# B&R Automation Studio project Palletizer_Final_project_2
Automation Studio 4.10.2.37

## Configuration Config1

### Hardware
```
4PP065_0351_P74 : 4PP065.0351-P74 v1.0.4.0
  Connector IF5:
    ActivateDevice = 1
    Mode = Manual
    InternetAddress = 127.0.0.1
    Vnc1
    VncVcObjectName1 = Visu_R
    VncKeyMappingFile1 = VC\PS2-Keyboard.dis
    VncAuthentication1 = 1
    VncPasswordViewOnly1 = r
    VncPasswordViewControl1 = w
  ConfigurationID = Palletizer_Final_project_Config1
  Simulation = 1
  FileDevice1
  FileDeviceName1 = USER
  FileDevicePath1 = USER_PATH
  KeyMappingFile = VC\4PP065_0351_P74.dis
```

## Logical view

Binary libraries used (declarations not repeated): operator, runtime, astime, AsIecCon, AsTCP, standard, AsArLog, AsBrStr

### Global.var - Global variables
```iecst
(*FEEDERSTATION*)
(*Insert your comment here.*)
VAR
	OperationType : INT;
	ENABLE_CONVEYER_END : BOOL;
	ENABLE_CONVEYER_TURN1 : BOOL;
	TURNPUSHER_FAULT : BOOL;
	ENABLE_TURNPUSHER : BOOL;
	DISABLE_TURNPUSHER : BOOL;
	TURNPUSHER_ENABLED : BOOL;
	TURNPUSHER_DISABLED : BOOL;
	PUSHER_FAULT : BOOL;
	ENABLE_PUSHER : BOOL;
	PUSHER_DISABLED : BOOL;
	PUSHER_ENABLED : BOOL;
	ENABLE_CONVEYOR_IF : BOOL;
	START_FEEDER : BOOL;
	LASER_SENSOR_IR : BOOL;
	FIRST_LAYER_OPERATION : BOOL;
	NUM_BOX_COUNTED : INT;
	COUNT_LASER_SENSOR_IR : INT;
	LASER_SENSOR_2_IR : BOOL;
	ACTUAL_BOXES : INT;
	ACTUAL_CARRIAGE_POS : REAL;
	CARRIAGE_TRG_POS : REAL;
	CARRIAGE_RCHD_POS : BOOL;
	SIMULATE_FAULT_CARRIAGE_2 : BOOL;
	FEERDER_BOXES_DELIVERED : BOOL;
	START_AGAIN_FEEDER : BOOL;
	FEEDER_EMERGENCY_STOP : BOOL;
	FEEDER_IMMEDIATE_STOP : BOOL;
	FEEDER_ON_PHASE_STOP : BOOL;
	FEEDER_ON_PHASE_STOP_WAIT : BOOL;
	ENABLE_SLIDE_RAIL_RIGHT : BOOL;
	VACUUM_BOX_CRANE_ENABLED : BOOL;
	ENABLE_VACUUM_BOX_CRANE : BOOL;
	VACUUM_BOX_CRANE_FAULT : BOOL;
	ENABLE_PUSHER_X : BOOL;
	ENABLE_PUSHER_Z : BOOL;
	ENABLE_CARTBORAD : BOOL;
	GANTRY_CRANE_RCHD_POS : BOOL;
	FAULT_GANTRY_CRANE : BOOL;
	ACTUAL_GANTRY_CRANE_POS : REAL;
	GANTRY_CRANE_TRG_POS : REAL;
	BOX_CRANE_RCHD_POS : BOOL;
	FAULT_BOX_CRANE : BOOL;
	ACTUAL_BOX_CRANE_POS : REAL;
	BOX_CRANE_TRG_POS : REAL;
	START_CRANE : BOOL;
	CRANE_WAIT_BOXES : BOOL;
	SECOND_LAYER_OPERATION : BOOL;
	LASER_SENSOR_IR_MEM : BOOL;
	LASER_SENSOR_2_IR_MEM : BOOL;
	CRANE_ON_PHASE_STOP : BOOL;
	CRANE_ON_PHASE_STOP_WAIT : BOOL;
	CRANE_EMERGENCY_STOP : BOOL;
	CRANE_IMMEDIATE_STOP : BOOL;
	FAULT_PALLET_CONVEYOR_2 : BOOL;
	PALLET_CONVEYOR_2_TRG_VEL : REAL;
	PALLET_LIFTER_RCHD_POS : BOOL;
	FAULT_PALLET_LIFTER : BOOL;
	ACTUAL_PALLET_LIFTER_POS : REAL;
	PALLET_LIFTER_TRG_POS : REAL;
	PALLET_FORK_ENABLED : BOOL;
	ENABLE_PALLET_FORK : BOOL;
	PALLET_FORK_FAULT : BOOL;
	ENABLE_PALLET_CONVEYOR_1 : BOOL;
	PALLET_CONVEYOR_1_FAULT : BOOL;
	PALLET_LIGHT_BARRIER_2 : BOOL;
	PALLET_LIGHT_BARRIER_1 : BOOL;
	PALLET_WAIT_BOXES : BOOL;
	AFTER_IMMEDIATE_STOP : BOOL; (*gives acces to the pallet state after the immediate stop*)
	START_PALLET : BOOL;
	PALLET_ON_PHASE_STOP_WAIT : BOOL;
	PALLET_EMERGENCY_STOP : BOOL;
	PALLET_IMMEDIATE_STOP : BOOL;
	PALLET_ON_PHASE_STOP : BOOL;
	BUTTON_START : BOOL;
	BUTTON_STOP : BOOL;
	BUTTON_EMERGENCY_STOP : BOOL;
	BUTTON_IMMEDIATE_STOP : BOOL;
	BUTTON_ON_PHASE_STOP : BOOL;
	BUTTON_INITIALIZATION : BOOL;
	blink_start : BOOL;
	blink_stop : BOOL;
	blink_ermergency : BOOL;
	blink_immediatestop : BOOL;
	blink_onphasestop : BOOL;
	blink_Fauld : BOOL;
	FEERDER_WAIT_TO_DELIVER_BOXES : BOOL;
	CRANE_BOXES_DELIVERED : BOOL;
	CARRIAGE_2_FAULT : BOOL;
	CONVEYOR_IF_FAULT : BOOL;
	SIMULATE_FAULT_PUSHER : BOOL;
	SIMULATE_FAULT_TURNPUSHER : BOOL;
	SIMULATE_FAULT_GANTRY_CRANE : BOOL;
	GANTRY_CRANE_FAULT : BOOL;
	SIMULATE_FAULT_BOX_CRANE : BOOL;
	BOX_CRANE_FAULT : BOOL;
	SIMULATE_FAULT_SLIDE_RIGTH : BOOL;
	SIMULATE_FAULT_SLIDE_RAIL_RIGHT : BOOL;
	SLIDE_RAIL_RIGHT_FAULT : BOOL;
	SIMULATE_FAULT_VACUUM_BOX_CRANE : BOOL;
	SIMULATE_FAULT_PUSHER_X : BOOL;
	PUSHER_X_FAULT : BOOL;
	SIMULATE_FAULT_PUSHER_Z : BOOL;
	PUSHER_Z_FAULT : BOOL;
	SIMULATE_FAULT_CARTBORAD : BOOL;
	CARTBORAD_FAULT : BOOL;
	SIMULATE_FAULT_PALLET_LIFTER : BOOL;
	PALLET_LIFTER_FAULT : BOOL;
	SIMULATE_FAULT_PALLET_CONVEYOR_2 : BOOL;
	PALLET_CONVEYOR_2_FAULT : BOOL;
	SIMULATE_FAULT_PALLET_FORK : BOOL;
	ENABLE_CONVEYOR_TURN1 : BOOL;
	CONVEYOR_TURN1_FAULT : BOOL;
	ENABLE_CONVEYOR_END : BOOL;
	CONVEYOR_END_FAULT : BOOL;
	LED_ALARM_INFORMATION : BOOL;
	LED_ALARM_ANOMALY : BOOL;
	LED_ALARM_ALARM : BOOL;
	LED_ALARM_WARNING : BOOL;
	SM_ON_PHASE_STOP : BOOL;
	SM_IMMEDIATE_STOP : BOOL;
	SM_EMERGENCY_STOP : BOOL;
	SM_IMMEDIATE_STOP_CAT1 : BOOL;
	SM_IMMEDIATE_STOP_CAT2 : BOOL;
	SM_IMMEDIATE_STOP_CAT3 : BOOL;
	LED_MATERIALS_RUN_OUT : BOOL;
	SM_ON_PHASE_STOP_CAT2 : BOOL;
	SM_ON_PHASE_STOP_CAT1 : BOOL;
	PALLET_ON_PHASE_STOP_REMOVE : BOOL;
	SM_ON_PHASE_STOP_CAT_2 : BOOL;
	boxcrane_Cartboard_ALMOST_FINISH : BOOL;
	boxcrane_Cartboard_FINISH : BOOL;
	pallet_lifter_ALMOST_FINISH : BOOL;
	pallet_lifter_FINISH : BOOL;
	POWER_ON_FEEDER : BOOL;
	POWER_ON_CRANE : BOOL;
	POWER_ON_PALLET : BOOL;
	POWER_MACHINE : BOOL;
	POWER_ON_BUTTON : BOOL;
	PALLET_ON_PHASE_STOP_IDLE : BOOL;
	COUNT_PALLET_NUMBER : INT := 5;
	COUNT_CARTBOARD_NUMBER : INT := 25;
	COUNT_BOXES_NUMBER : INT;
	blink_emergencvy_stop : BOOL;
	blink_immediate_stop : BOOL;
	blink_OnPhase_stop : BOOL;
	PALLET_STOP : BOOL;
	CRANE_STOP : BOOL;
	FEEDER_STOP : BOOL;
END_VAR
```

### MNG_Package.var
```iecst
(*                                                                            *)
(* File generated by the B&R AS 4 control config generator                    *)
(*                                                                            *)
(*     Provider: machineering                                                 *)
(*  Application: industrialPhysics_2.4.master                                 *)
(* Architecture: Windows 64 Bit                                               *)
(*      Version: 2.4.10491.master                                             *)
(*        Build: 164f85bec                                                    *)
(*         Date: 2020-05-19, Time: 12:11:21                                   *)
(*                                                                            *)
VAR
	ComTCP_SimInputs : ComTCP_INPUTS_32BIT := (0);
	ComTCP_SimOutputs : ComTCP_OUTPUTS_32BIT := (0);
	ComTCP_SimServerAddress : STRING[15] := '127.0.0.1';
	ComTCP_SimServerPort : UINT := 5000;
	ComTCP_SimSendCycleTime : TIME := T#5ms;
	ComTCP_SimActive : BOOL := FALSE;
END_VAR
```

### MNG_Package.typ
```iecst
(*                                                                            *)
(* File generated by the B&R AS 4 control config generator                    *)
(*                                                                            *)
(*     Provider: machineering                                                 *)
(*  Application: industrialPhysics_2.4.master                                 *)
(* Architecture: Windows 64 Bit                                               *)
(*      Version: 2.4.10491.master                                             *)
(*        Build: 164f85bec                                                    *)
(*         Date: 2020-05-19, Time: 12:11:21                                   *)
(*                                                                            *)

TYPE
	ComTCP_INPUTS_32BIT : 	STRUCT
		NumSignals : INT := 15;
		laser_sensor_IR : BOOL := 0; (* BOOL laser_sensor_IR *)
		laser_sensor2_IR : BOOL := 0; (* BOOL laser_sensor2_IR *)
		carriage_2_AXIS : REAL := 0.0; (* REAL carriage_2_AXIS *)
		carriage_2_RCHD : BOOL := 0; (* BOOL carriage_2_RCHD *)
		turnpusher_LBK : BOOL := 0; (* BOOL turnpusher_LBK *)
		turnpusher_LFR : BOOL := 0; (* BOOL turnpusher_LFR *)
		gantry_crane_AXIS : REAL := 0.0; (* REAL gantry_crane_AXIS *)
		box_crane_AXIS : REAL := 0.0; (* REAL box_crane_AXIS *)
		vaccum_box_crane_VACUUM : BOOL := 0; (* BOOL vaccum_box_crane_VACUUM *)
		pallet_light_barrier_1_IR : BOOL := 0; (* BOOL pallet_light_barrier_1_IR *)
		pallet_light_barrier_2_IR : BOOL := 0; (* BOOL pallet_light_barrier_2_IR *)
		pusher_LBK : BOOL := 0; (* BOOL pusher_LBK *)
		pusher_LFR : BOOL := 0; (* BOOL pusher_LFR *)
		pallet_lifter_AXIS : REAL := 0.0; (* REAL pallet_lifter_AXIS *)
		pallet_fork_left_FB : BOOL := 0; (* BOOL pallet_fork_left_FB *)
	END_STRUCT;
	ComTCP_OUTPUTS_32BIT : 	STRUCT
		NumSignals : INT := 18;
		cartboard_TRIG : BOOL := 0; (* BOOL cartboard_TRIG *)
		conveyor_if_FWD : BOOL := 0; (* BOOL conveyor_if_FWD *)
		conveyer_turn1_FWD : BOOL := 0; (* BOOL conveyer_turn1_FWD *)
		conveyer_end_FWD : BOOL := 0; (* BOOL conveyer_end_FWD *)
		carriage_2_TGT_POS : REAL := 0.0; (* REAL carriage_2_TGT_POS *)
		turnpusher_FWD : BOOL := 0; (* BOOL turnpusher_FWD *)
		turnpusher_BWD : BOOL := 0; (* BOOL turnpusher_BWD *)
		gantry_crane_TGT_POS : REAL := 0.0; (* REAL gantry_crane_TGT_POS *)
		box_crane_TGT_POS : REAL := 0.0; (* REAL box_crane_TGT_POS *)
		slide_rail_right_EN : BOOL := 0; (* BOOL slide_rail_right_EN *)
		vaccum_box_crane_GRIP : BOOL := 0; (* BOOL vaccum_box_crane_GRIP *)
		pusher_z_EN : BOOL := 0; (* BOOL pusher_z_EN *)
		pusher_x_EN : BOOL := 0; (* BOOL pusher_x_EN *)
		pallet_conveyor_2_ACT_VEL : REAL := 0.0; (* REAL pallet_conveyor_2_ACT_VEL *)
		pusher_FW : BOOL := 0; (* BOOL pusher_FW *)
		pallet_lifter_TGT_POS : REAL := 0.0; (* REAL pallet_lifter_TGT_POS *)
		pallet_fork_left_EN : BOOL := 0; (* BOOL pallet_fork_left_EN *)
		pallet_conveyor_1_FWD : BOOL := 0; (* BOOL pallet_conveyor_1_FWD *)
	END_STRUCT;
END_TYPE
```

### Package Logical/Libraries - Global libraries

### Library Logical/Libraries/G_Device (IEC)

#### Types.typ - Exported data types
```iecst
TYPE
	DeviceStateType :
	(
		DeviceEnabledState		:=2,
		DeviceEnablePhaseState	:=1,
		DeviceDisabledState		:=0,
		DeviceDisablePhaseState	:=3
	);
END_TYPE
```

#### Constants.var - Exported constants
```iecst
VAR CONSTANT
	DEVICE_ACTUATION_MASK : INT := 2#00001111;
	DEVICE_FEEDBACK_MASK : INT := 2#11110000;
	DEVICE_WITH_ENABLE_FEEDBACK : INT := 2#00010000;
	DEVICE_WITH_DISABLE_FEEDBACK : INT := 2#00100000;
	DEVICE_WITHOUT_FEEDBACK : INT := 2#01000000;
	DEVICE_WITH_SINGLE_ACTUATION : INT := 2#00000001;
	DEVICE_WITH_DOUBLE_ACTUATION : INT := 2#00000011;
	DEVICE_WITH_DA_NO_RETAIN : INT := 2#00000010;
	DEVICE_WITH_DOUBLE_FEEDBACK : INT := 2#00110000;
END_VAR
```

#### G_Device.fun - Exported functions and function blocks
```iecst
{REDUND_ERROR} FUNCTION_BLOCK Generic_Device (*TODO: Add your comment here*) (*$GROUP=User,$CAT=User,$GROUPICON=User.png,$CATICON=User.png*)
	VAR_INPUT
		DeviceClock : {REDUND_UNREPLICABLE} BOOL;
		DeviceDisabledSensor : {REDUND_UNREPLICABLE} BOOL;
		DeviceEnabledSensor : {REDUND_UNREPLICABLE} BOOL;
		DeviceEnabled : {REDUND_UNREPLICABLE} BOOL;
		DeviceDisabled : {REDUND_UNREPLICABLE} BOOL;
		DeviceType : {REDUND_UNREPLICABLE} INT;
		DeviceOperation : {REDUND_UNREPLICABLE} INT;
		DeviceEnablePreset : {REDUND_UNREPLICABLE} BOOL;
		DeviceEnableTime : {REDUND_UNREPLICABLE} INT;
		DeviceDisableTime : {REDUND_UNREPLICABLE} INT;
		DeviceDiagnosticsEnabled : BOOL;
		SimulationDeviceFault : BOOL;
	END_VAR
	VAR_OUTPUT
		EnableDevice : {REDUND_UNREPLICABLE} BOOL;
		DeviceNotInitialized : {REDUND_UNREPLICABLE} BOOL;
		DisableDevice : {REDUND_UNREPLICABLE} BOOL;
		DeviceDisabledSensorFault : {REDUND_UNREPLICABLE} BOOL;
		DeviceEnabledSensorFault : {REDUND_UNREPLICABLE} BOOL;
		DeviceActuatorFault : {REDUND_UNREPLICABLE} BOOL;
		DeviceFault : {REDUND_UNREPLICABLE} BOOL;
	END_VAR
	VAR_IN_OUT
		DeviceEnableRequest : BOOL;
		DeviceDisableRequest : BOOL;
	END_VAR
	VAR
		DeviceTimer : {REDUND_UNREPLICABLE} INT;
	END_VAR
	VAR RETAIN
		DeviceState : {REDUND_UNREPLICABLE} DeviceStateType;
	END_VAR
	VAR
		Timeout : {REDUND_UNREPLICABLE} BOOL := FALSE;
	END_VAR
	VAR CONSTANT
		INIT : INT := 0;
	END_VAR
	VAR
		WaitNominalStateCounter : INT := 20;
		SimulationDeviceActuatorFault : BOOL;
	END_VAR
END_FUNCTION_BLOCK
```

#### Generic_Device.st
```iecst
(* TODO: Add your comment here *)
FUNCTION_BLOCK Generic_Device

	//I-) DEVICE CLOCK HANDLER
	IF (DeviceClock AND (DeviceTimer > 0))THEN
		DeviceTimer := DeviceTimer - 1;
		WaitNominalStateCounter := WaitNominalStateCounter	- 1;
	END_IF;

	//II-) DEVICE SENSORS HANDLER
	CASE (DeviceType AND DEVICE_FEEDBACK_MASK) OF

		DEVICE_WITH_ENABLE_FEEDBACK:

			DeviceDisabledSensor := NOT DeviceEnabledSensor AND
			((DeviceState = DeviceDisabledState) OR (DeviceState = DeviceDisablePhaseState AND Timeout));
			//Pre-elaborations actuators
			DeviceDisabled := NOT DeviceEnabled AND ((DeviceState = DeviceDisabledState) OR
			(DeviceState = DeviceDisablePhaseState AND Timeout));

		DEVICE_WITH_DISABLE_FEEDBACK :

			DeviceEnabledSensor := NOT DeviceDisabledSensor AND
			((DeviceState = DeviceEnabledState) OR (DeviceState = DeviceEnablePhaseState AND Timeout));
			//Pre-elaborations actuators
			DeviceEnabled := NOT DeviceDisabled AND ((DeviceState = DeviceEnabledState) OR
			(DeviceState = DeviceEnablePhaseState AND Timeout));

		DEVICE_WITHOUT_FEEDBACK:

			DeviceEnabledSensor := (DeviceState = DeviceEnabledState) OR ((DeviceState = DeviceEnablePhaseState) AND Timeout);
			DeviceDisabledSensor := (DeviceState = DeviceDisabledState) OR ((DeviceState = DeviceDisablePhaseState) AND Timeout);
			//Pre-elaborations actuators
			DeviceEnabled := (DeviceState = DeviceEnabledState) OR (DeviceState = DeviceEnablePhaseState AND Timeout);
			DeviceDisabled := (DeviceState = DeviceDisabledState) OR (DeviceState = DeviceDisablePhaseState AND Timeout);

	END_CASE;

	//III-) DEVICE INITIALIZATION HANDLER
	IF (DeviceOperation = INIT) THEN
		// Device sensor handler
		CASE (DeviceType AND DEVICE_FEEDBACK_MASK) OF

			DEVICE_WITH_ENABLE_FEEDBACK:
				DeviceDisabled := NOT DeviceEnabled;

			DEVICE_WITH_DISABLE_FEEDBACK :
				DeviceEnabled := NOT DeviceDisabled;

			DEVICE_WITHOUT_FEEDBACK:
				DeviceEnabled := DeviceEnablePreset;
				DeviceDisabled := NOT DeviceEnabled;

		END_CASE;

		DeviceEnableRequest := FALSE;
		DeviceDisableRequest := FALSE;

		IF (DeviceEnablePreset) THEN
			EnableDevice := TRUE;
			DeviceTimer := DeviceEnableTime;
			IF (NOT (DeviceDisabled AND DeviceEnabled)) THEN
				DeviceState := DeviceEnablePhaseState;
			ELSE
				DeviceState := DeviceEnabledState;
			END_IF;
			DeviceNotInitialized := NOT DeviceEnabled OR DeviceDisabled;
		ELSE
			EnableDevice := FALSE;
			DeviceTimer := DeviceDisableTime;
			IF (NOT (DeviceDisabled AND DeviceEnabled)) THEN
				DeviceState := DeviceDisablePhaseState;
			ELSE
				DeviceState := DeviceDisabledState;
			END_IF;
			DeviceNotInitialized := (DeviceEnabled OR NOT DeviceDisabled);
		END_IF;
	END_IF;

	IF NOT SimulationDeviceFault THEN
		//IV-) DEVICE CONTROL HANDLER (GENERIC DEVICE FSM IMPLEMENTATION)
		CASE (DeviceState) OF

			DeviceDisabledState:
				DeviceDisableRequest := FALSE;
				IF (DeviceEnableRequest) THEN
					EnableDevice := TRUE;
					DeviceTimer := DeviceEnableTime;
					DeviceState := DeviceEnablePhaseState;
				END_IF;

			DeviceEnablePhaseState:
				IF DeviceDisableRequest THEN
					DeviceEnableRequest	:= FALSE;
					EnableDevice	:= FALSE;
					DeviceTimer	:= DeviceDisableTime;
					DeviceState	:= DeviceDisablePhaseState;
				END_IF;
				IF DeviceEnabledSensor THEN
					DeviceEnableRequest := FALSE;
					DeviceTimer	:= 0;
					DeviceState := DeviceEnabledState;
				END_IF;

			DeviceEnabledState:
				DeviceEnableRequest	:= FALSE;
				IF DeviceDisableRequest THEN
					EnableDevice := FALSE;
					DeviceTimer	:= DeviceDisableTime;
					DeviceState := DeviceDisablePhaseState;
				END_IF;

			DeviceDisablePhaseState:
				IF DeviceEnableRequest THEN
					DeviceDisableRequest	:= FALSE;
					EnableDevice	:= TRUE;
					DeviceTimer	:= DeviceEnableTime;
					DeviceState	:= DeviceEnablePhaseState;
				END_IF;

				IF DeviceDisabledSensor THEN
					DeviceDisableRequest := FALSE;
					DeviceTimer	:= 0;
					DeviceState := DeviceDisabledState;
				END_IF;

		END_CASE;

	END_IF;

	//handler timer
	IF (DeviceTimer = 0) THEN
		Timeout := TRUE ;

	ELSE
		Timeout := FALSE ;

	END_IF;

	//V-) DEVICE DIAGNOSTICS HANDLER (GENERATION OF DIAGNOSIS INFORMATION),
	DeviceDisabledSensorFault := (( NOT EnableDevice AND NOT DeviceDisabledSensor AND NOT DeviceEnabledSensor) OR (EnableDevice AND DeviceDisabledSensor AND DeviceEnabledSensor)) AND Timeout;

	DeviceEnabledSensorFault := ((NOT EnableDevice AND DeviceDisabledSensor AND DeviceEnabledSensor) OR (EnableDevice AND NOT DeviceDisabledSensor AND NOT DeviceEnabledSensor)) AND Timeout;

	DeviceActuatorFault := ((NOT EnableDevice AND NOT DeviceDisabledSensor AND DeviceEnabledSensor AND Timeout) OR (EnableDevice AND DeviceDisabledSensor AND NOT DeviceEnabledSensor AND Timeout)) AND Timeout;
	//DeviceActuatorFault

	DeviceFault :=	DeviceDisabledSensorFault OR DeviceEnabledSensorFault OR SimulationDeviceFault ;

	//VI-) DEVICE ACTUATORS HANDLER (Post-elaborations actustors)
	IF (DeviceType AND DEVICE_ACTUATION_MASK)= DEVICE_WITH_SINGLE_ACTUATION THEN
		//Nothing to do, just use EnableDevice
	END_IF;
	IF	(DeviceType AND DEVICE_ACTUATION_MASK)= DEVICE_WITH_DOUBLE_ACTUATION THEN
		DisableDevice := NOT EnableDevice;
	END_IF;
	IF	(DeviceType AND DEVICE_ACTUATION_MASK)= DEVICE_WITH_DA_NO_RETAIN THEN
		EnableDevice := EnableDevice AND (DeviceState = DeviceEnablePhaseState);
		DisableDevice := NOT EnableDevice AND (DeviceState = DeviceDisablePhaseState);
	END_IF;
	IF	DeviceActuatorFault AND (DeviceTimer = 0) AND WaitNominalStateCounter = 0  THEN

		SimulationDeviceActuatorFault := TRUE;
		WaitNominalStateCounter := 20;

	ELSE
		SimulationDeviceActuatorFault := FALSE;
	END_IF;

END_FUNCTION_BLOCK
```

### Library Logical/Libraries/G_Axis (IEC)

#### Types.typ - Exported data types
```iecst
TYPE

	GenericAxisType :
		(
		WaitpowerON,
		WaitHoming,
		CheckCommand,
		WaitPowerOFF,
		WaitStop,
		WaitMoveTRG_POS,
		ErrorState,
		WaitMoveTRG_VEL

	);

END_TYPE
```

#### Constants.var - Exported constants
```iecst
VAR CONSTANT
	POWEROFF : DWORD := 1;
	STOP : DWORD := 2;
	HOMING : DWORD := 3;
	TARGETPOSITION : DWORD := 4;
	Notbusy : DWORD := 0;
	TARGETVELOCITY : DWORD := 5;
END_VAR
```

#### G_Axis.fun - Exported functions and function blocks
```iecst
{REDUND_ERROR} FUNCTION_BLOCK Generic_Axis (*TODO: Add your comment here*) (*$GROUP=User,$CAT=User,$GROUPICON=User.png,$CATICON=User.png*)
	VAR_INPUT
		PowerON : BOOL;
		DeviceTimer : INT;
		Actual_position : REAL;
		Input_Target_Position : REAL;
		Reached_Postion : BOOL;
		InputSimulateError : BOOL;
		Actual_Command : DWORD;
		DeviceClock : BOOL;
		DeviceFeedback : BOOL;
	END_VAR
	VAR_OUTPUT
		Powered : BOOL;
		Output_Target_Position : REAL;
		InPosition : BOOL;
		InVelocity : BOOL;
		OutputSimulateError : BOOL;
	END_VAR
	VAR
		Generic_Axis_State : GenericAxisType;
		Timer : INT;
		TimeOut : BOOL;
	END_VAR
	VAR_INPUT
		Input_Target_Velocity : REAL;
	END_VAR
	VAR_OUTPUT
		Output_Target_Velocity : REAL;
	END_VAR
END_FUNCTION_BLOCK
```

#### Generic_Axis.st
```iecst
(* TODO: Add your comment here *)
FUNCTION_BLOCK Generic_Axis
	IF (DeviceClock AND (Timer > 0))THEN
		Timer := Timer - 1;

		END_IF;

	CASE Generic_Axis_State OF

		WaitpowerON:
			IF PowerON THEN
				//all output false
				Powered:= FALSE;
				InPosition	:= FALSE;
				InVelocity	:= FALSE;
				Timer		:= DeviceTimer;
	  			Generic_Axis_State:=WaitHoming;
			END_IF;
		WaitHoming:

			IF TimeOut THEN
				Powered:= TRUE;
				TimeOut		:= FALSE;
				Output_Target_Position:=0.0;
				Output_Target_Velocity:=0.0;
				Actual_Command := Notbusy;
				IF NOT PowerON THEN
					Generic_Axis_State:= WaitpowerON;
				ELSE
					IF Actual_position=0.0 THEN
						InPosition	:= TRUE;
						InVelocity	:= FALSE;
						Generic_Axis_State:= CheckCommand;
					END_IF;
				END_IF;
			END_IF;
		CheckCommand:
			IF Actual_Command = POWEROFF  THEN
				Actual_Command := Notbusy;
				Generic_Axis_State:= WaitPowerOFF;
			END_IF;
			IF Actual_Command = STOP THEN
				Actual_Command := Notbusy;
				Generic_Axis_State:= WaitStop;
			END_IF;
			IF Actual_Command = HOMING THEN
				Actual_Command := Notbusy;
				InVelocity	:= TRUE;
				Generic_Axis_State:= WaitHoming;
			END_IF;
			IF Actual_Command = TARGETPOSITION THEN
				Actual_Command := Notbusy;
				IF Input_Target_Position <> Actual_position THEN
					InVelocity	:= TRUE;
					Timer		:= DeviceTimer;
	  				Generic_Axis_State:= WaitMoveTRG_POS;
				ELSE
					Generic_Axis_State:= CheckCommand;
				END_IF;
			END_IF;
			InPosition	:= FALSE;
			IF Actual_Command = TARGETVELOCITY THEN
				Actual_Command := Notbusy;
				IF Input_Target_Velocity <> Output_Target_Velocity THEN
					InVelocity	:= TRUE;
					Timer		:= DeviceTimer;
					Generic_Axis_State:= WaitMoveTRG_VEL;
				ELSE
					Generic_Axis_State:= CheckCommand;
				END_IF;
			END_IF;
		WaitPowerOFF:
			PowerON := FALSE;
			InPosition	:= FALSE;
			InVelocity	:= FALSE;
			Generic_Axis_State:=WaitHoming;
		WaitStop:

			IF InVelocity THEN
		  		Output_Target_Position:=Actual_position + 0.1; //bias link to the dealy
				IF Reached_Postion THEN

		  			InPosition	:= FALSE;
					InVelocity	:= FALSE;
				END_IF;
			END_IF;
			IF OutputSimulateError THEN
				Generic_Axis_State:= ErrorState;
			ELSE
				Generic_Axis_State:= CheckCommand;
			END_IF;

		WaitMoveTRG_POS:
			Output_Target_Position := Input_Target_Position;
			IF TimeOut THEN
				IF DeviceFeedback AND Reached_Postion THEN
					InPosition	:= TRUE;
					InVelocity	:= FALSE;
					TimeOut		:= FALSE;
					Generic_Axis_State:= CheckCommand;
				END_IF;

				IF NOT DeviceFeedback AND (Input_Target_Position = Actual_position)	 THEN
					InPosition	:= TRUE;
					InVelocity	:= FALSE;
					TimeOut		:= FALSE;
					Generic_Axis_State:= CheckCommand;
				END_IF;

			END_IF;
		WaitMoveTRG_VEL:
			Output_Target_Velocity := Input_Target_Velocity;
			IF TimeOut THEN
				IF NOT DeviceFeedback THEN
					TimeOut		:= FALSE;
					Generic_Axis_State:= CheckCommand;
				END_IF;
			END_IF;

		ErrorState:
			IF NOT InputSimulateError THEN //wait for the Simulated Error to be set back
				OutputSimulateError:=FALSE;
			Generic_Axis_State:= WaitHoming;
			END_IF;

	END_CASE;
	IF Timer=0 THEN
		TimeOut	:= TRUE;
	END_IF;
	IF InputSimulateError THEN
		OutputSimulateError:=TRUE;
		Generic_Axis_State:= WaitStop;
	END_IF;

END_FUNCTION_BLOCK
```

### Library Logical/Libraries/G_SM (IEC)

#### Constants.var - Exported constants
```iecst
VAR CONSTANT
	SIGNAL_TYPE_MASK : INT := 2#00000111;
	ALARM : INT := 2#00000001;
	ANOMALY : INT := 2#00000010;
	WARNING : INT := 2#00000011;
	INFORMATION : INT := 2#00000100;
	AUX_RESET : INT := 2#10100000;
	AUTO_CONDITIONED_RESET : INT := 2#01100000;
	NONE : DWORD := 16#0000;
	INIT : INT := 0;
	RUN : INT := 1;
	START_CONFIGURATION : INT := 2;
	CONFIGURATION : INT := 3;
	START_GENERATION : INT := 4;
	GENERATION : INT := 5;
	EMERGENCY_STOP : DWORD := 16#0001;
	IMMEDIATE_STOP : DWORD := 16#0002;
	ON_PHASE_STOP : DWORD := 16#0004;
	MATERIALS_RUN_OUT_LAMP : DWORD := 16#0006;
	MATERIALS_RUN_OUT_BUZZER : DWORD := 16#0008;
END_VAR
```

#### G_SM.fun - Exported functions and function blocks
```iecst
{REDUND_ERROR} FUNCTION_BLOCK GenericSignalHandler (*TODO: Add your comment here*) (*$GROUP=User,$CAT=User,$GROUPICON=User.png,$CATICON=User.png*)
	VAR_INPUT
		OperationType : INT;
		SignalType : DINT;
		Reset : BOOL;
		KeyReset : BOOL;
		ActivationSignal : BOOL;
		SignalCode : INT;
		SignalOutput : DWORD;
		CondKeyReset : BOOL;
	END_VAR
	VAR_OUTPUT
		NumberOfAlarms : INT;
		NumberOfAnomalies : INT;
		NumberOfWarnings : INT;
		NumberOfInformation : INT;
		ResetEnable : BOOL;
		SignalOutputs : DWORD;
		NumberOfActiveAlarms : INT;
		NumberOfActiveAnomalies : INT := 0;
		NumberOfActiveWarning : INT;
		NumberOfActiveInformation : INT;
		ActiveSignalCodes : ARRAY[0..24] OF INT;
		AuxResetEnable : BOOL;
		AutoCondResetEnable : BOOL;
		LedSignalInformation : BOOL;
		LedSignalAnomaly : BOOL;
		LedSignalWarning : BOOL;
		LedSignalAlarm : BOOL;
		MySignalCode : INT;
	END_VAR
	VAR
		ResetActivation : BOOL;
		ResetOld : BOOL;
		KeyResetOld : BOOL;
		Index : INT;
		BaseIndex : INT;
		Condition : BOOL;
		Signals : {REDUND_UNREPLICABLE} ARRAY[0..24] OF BOOL;
		i : INT;
		AuxResetActivation : BOOL;
		AuxResetOfSignalType : BOOL;
		AutoCondResetOfSignalType : BOOL;
		AutoCondResetActivation : BOOL;
		CondKeyResetOld : BOOL;
	END_VAR
END_FUNCTION_BLOCK
```

#### GenericSignalHandler.st
```iecst
(* TODO: Add your comment here *)
FUNCTION_BLOCK GenericSignalHandler

	CASE OperationType OF

		INIT:

		START_CONFIGURATION: (* Reset signals counts *)

			NumberOfAlarms := 0;
			NumberOfAnomalies := 0;
			NumberOfWarnings := 0;
			NumberOfInformation := 0;

		CONFIGURATION: (* counting signals *)

			CASE (SignalType AND SIGNAL_TYPE_MASK) OF
				ALARM:
					NumberOfAlarms := NumberOfAlarms + 1;
				ANOMALY:
					NumberOfAnomalies := NumberOfAnomalies + 1;
				WARNING:
					NumberOfWarnings := NumberOfWarnings + 1;
				INFORMATION:
					NumberOfInformation := NumberOfInformation + 1;
			END_CASE

		START_GENERATION: (* Prepare for generation *)

			ResetEnable := FALSE;
			SignalOutputs := NONE;
			ResetActivation := Reset AND NOT ResetOld;
			ResetOld := Reset;
			AuxResetActivation := KeyReset AND NOT KeyResetOld;
			KeyResetOld := KeyReset;
			AutoCondResetActivation := CondKeyReset AND NOT CondKeyResetOld;

			CondKeyResetOld := CondKeyReset;
		GENERATION:
			CASE (SignalType AND SIGNAL_TYPE_MASK) OF
				ALARM:
					Index := NumberOfActiveAlarms;
					BaseIndex := 0;
					Condition := TRUE;
				ANOMALY:
					Index := NumberOfActiveAnomalies;
					BaseIndex := NumberOfAlarms;
					Condition := TRUE;
				WARNING:
					Index := NumberOfActiveWarning;
					BaseIndex := NumberOfAlarms + NumberOfAnomalies;
					Condition := FALSE;
				INFORMATION:
					Index := NumberOfActiveInformation;
					BaseIndex := NumberOfAlarms + NumberOfAnomalies + NumberOfWarnings;
					Condition := FALSE;
			END_CASE

			IF ActivationSignal AND NOT Signals[SignalCode] THEN
				Signals[SignalCode] := TRUE;
				Index := Index + 1;
				ActiveSignalCodes[BaseIndex + Index] := SignalCode;
			END_IF

			// Autoconditioned reset
			AutoCondResetOfSignalType := ((SignalType AND AUTO_CONDITIONED_RESET) = AUTO_CONDITIONED_RESET);

			IF Condition AND Signals[SignalCode] AND NOT ActivationSignal AND (ActiveSignalCodes[BaseIndex + 1] = SignalCode) AND AutoCondResetOfSignalType THEN
				AutoCondResetEnable := TRUE;

			END_IF

			// Auxiliary reset
			AuxResetOfSignalType := ((SignalType AND AUX_RESET) = AUX_RESET);
			IF Condition AND Signals[SignalCode] AND NOT ActivationSignal AND (ActiveSignalCodes[BaseIndex + 1] = SignalCode) AND AuxResetOfSignalType AND NOT AutoCondResetOfSignalType THEN
				AuxResetEnable := TRUE;

			END_IF

			//Direct reset
			IF Condition AND Signals[SignalCode] AND NOT ActivationSignal AND (ActiveSignalCodes[BaseIndex + 1] = SignalCode) AND NOT
				AuxResetOfSignalType  AND NOT AutoCondResetOfSignalType THEN
				ResetEnable := TRUE;
			END_IF

			IF (ResetActivation OR NOT Condition) AND Signals[SignalCode] AND NOT ActivationSignal AND
				(ActiveSignalCodes[BaseIndex + 1] = SignalCode)  AND NOT AutoCondResetOfSignalType AND NOT AuxResetOfSignalType THEN
				Signals[SignalCode] := FALSE;

				FOR i := 2 TO Index DO
					ActiveSignalCodes[BaseIndex + i-1] := ActiveSignalCodes[BaseIndex + i];
				END_FOR;
				ActiveSignalCodes[BaseIndex + Index] := 0;
				Index := Index - 1;
				ResetActivation := FALSE; (* COMMENT THIS LINE TO GO BACK TO CUMULATIVE RESET *)

			END_IF
			// Auxiliary reset
			IF (AuxResetActivation OR NOT Condition) AND Signals[SignalCode] AND NOT ActivationSignal AND
				(ActiveSignalCodes[BaseIndex + 1] = SignalCode) AND AuxResetOfSignalType  AND NOT AutoCondResetOfSignalType THEN
				Signals[SignalCode] := FALSE;

				FOR i := 2 TO Index DO
					ActiveSignalCodes[BaseIndex + i-1] := ActiveSignalCodes[BaseIndex + i];
				END_FOR;
				ActiveSignalCodes[BaseIndex + Index] := 0;
				Index := Index - 1;
				AuxResetActivation := FALSE; (* COMMENT THIS LINE TO GO BACK TO CUMULATIVE RESET *)

			END_IF
			// Autoconditioned reset
			IF (AutoCondResetActivation OR NOT Condition) AND Signals[SignalCode] AND NOT ActivationSignal AND
				(ActiveSignalCodes[BaseIndex + 1] = SignalCode) AND AuxResetOfSignalType AND AutoCondResetOfSignalType THEN
				Signals[SignalCode] := FALSE;

				FOR i := 2 TO Index DO
					ActiveSignalCodes[BaseIndex + i-1] := ActiveSignalCodes[BaseIndex + i];
				END_FOR;
				ActiveSignalCodes[BaseIndex + Index] := 0;
				Index := Index - 1;
				AutoCondResetActivation := FALSE; (* COMMENT THIS LINE TO GO BACK TO CUMULATIVE RESET *)

			END_IF

			CASE (SignalType AND SIGNAL_TYPE_MASK) OF
				ALARM:
					NumberOfActiveAlarms := Index;
				ANOMALY:
					NumberOfActiveAnomalies := Index;
				WARNING:
					NumberOfActiveWarning := Index;
				INFORMATION:
					NumberOfActiveInformation := Index;
			END_CASE
			IF Signals[SignalCode] THEN
				SignalOutputs := SignalOutputs OR SignalOutput;
				MySignalCode := SignalCode;

			END_IF

		RUN:
		(* UPDATE THE USER INTERFACE LED *)

			IF NumberOfActiveInformation >0 THEN

				LedSignalInformation	:= TRUE;

			ELSE
				LedSignalInformation	:= FALSE;
			END_IF

			IF NumberOfActiveAnomalies >0 THEN

				LedSignalAnomaly	:= TRUE;

			ELSE
				LedSignalAnomaly	:= FALSE;
			END_IF

			IF NumberOfActiveWarning >0 THEN

				LedSignalWarning	:= TRUE;

			ELSE
				LedSignalWarning	:= FALSE;
			END_IF

			IF NumberOfActiveAlarms >0 THEN

				LedSignalAlarm	:= TRUE;

			ELSE
				LedSignalAlarm	:= FALSE;
			END_IF

	END_CASE

END_FUNCTION_BLOCK
```

### Program Logical/Output_Bridge (IEC)

#### Main.st - Init, cyclic, exit code
```iecst
PROGRAM _INIT
	(* Insert code here *)

END_PROGRAM

PROGRAM _CYCLIC
	(* Insert code here *)
//CARRIAGE STATION
	ComTCP_SimOutputs.carriage_2_TGT_POS:=CARRIAGE_TRG_POS;

	ComTCP_SimOutputs.conveyor_if_FWD :=ENABLE_CONVEYOR_IF;
	ComTCP_SimOutputs.pusher_FW	:= ENABLE_PUSHER;
	ComTCP_SimOutputs.conveyer_turn1_FWD :=ENABLE_CONVEYOR_TURN1;
	ComTCP_SimOutputs.conveyer_end_FWD :=ENABLE_CONVEYOR_END;
	ComTCP_SimOutputs.turnpusher_FWD	:= DISABLE_TURNPUSHER;
	ComTCP_SimOutputs.turnpusher_BWD	:= ENABLE_TURNPUSHER;
//CRANE STATION
	ComTCP_SimOutputs.box_crane_TGT_POS		:= BOX_CRANE_TRG_POS;
	ComTCP_SimOutputs.cartboard_TRIG		:= ENABLE_CARTBORAD;
	ComTCP_SimOutputs.gantry_crane_TGT_POS	:= GANTRY_CRANE_TRG_POS;
	ComTCP_SimOutputs.pusher_x_EN			:= ENABLE_PUSHER_X;
	ComTCP_SimOutputs.pusher_z_EN			:= ENABLE_PUSHER_Z;
	ComTCP_SimOutputs.slide_rail_right_EN	:= ENABLE_SLIDE_RAIL_RIGHT;
	ComTCP_SimOutputs.vaccum_box_crane_GRIP	:= ENABLE_VACUUM_BOX_CRANE;
//PALLET STATION
	ComTCP_SimOutputs.pallet_lifter_TGT_POS	:= PALLET_LIFTER_TRG_POS;
	ComTCP_SimOutputs.pallet_fork_left_EN	:= ENABLE_PALLET_FORK;
	ComTCP_SimOutputs.pallet_conveyor_1_FWD	:= ENABLE_PALLET_CONVEYOR_1;
	ComTCP_SimOutputs.pallet_conveyor_2_ACT_VEL	:= PALLET_CONVEYOR_2_TRG_VEL;
	ComTCP_SimOutputs.pallet_lifter_TGT_POS	:= PALLET_LIFTER_TRG_POS;
//	ComTCP_SimOutputs.NumSignals
END_PROGRAM

PROGRAM _EXIT
	(* Insert code here *)

END_PROGRAM
```

#### Variables.var - Local variables
```iecst
VAR
	Activate_pusher_SA_SF : BOOL;
	Activate_turnpusher_DA_DF_FWD : BOOL;
	Activate_turnpusher_DA_DF_BWD : BOOL;
END_VAR
```

### Program Logical/Input_Bridge (IEC)

#### Main.st - Init, cyclic, exit code
```iecst
PROGRAM _INIT
	(* Insert code here *)

END_PROGRAM

PROGRAM _CYCLIC
	(* Insert code here *)
//CARRIAGE STATION
	LASER_SENSOR_2_IR	:= ComTCP_SimInputs.laser_sensor2_IR;
	LASER_SENSOR_IR		:= ComTCP_SimInputs.laser_sensor_IR;
	PUSHER_DISABLED		:= ComTCP_SimInputs.pusher_LBK ;
	PUSHER_ENABLED		:= ComTCP_SimInputs.pusher_LFR	;
	TURNPUSHER_DISABLED:= ComTCP_SimInputs.turnpusher_LBK;
	TURNPUSHER_ENABLED:= ComTCP_SimInputs.turnpusher_LFR;
	ACTUAL_CARRIAGE_POS := ComTCP_SimInputs.carriage_2_AXIS;
	CARRIAGE_RCHD_POS 	:= ComTCP_SimInputs.carriage_2_RCHD;
//	ComTCP_SimInputs.NumSignals

//CRANE STATION
	ACTUAL_BOX_CRANE_POS    := ComTCP_SimInputs.box_crane_AXIS;
	ACTUAL_GANTRY_CRANE_POS := ComTCP_SimInputs.gantry_crane_AXIS;
	VACUUM_BOX_CRANE_ENABLED:= ComTCP_SimInputs.vaccum_box_crane_VACUUM;

	(*INPUT FILTER*)
	IF LASER_SENSOR_IR THEN
		LASER_SENSOR_IR_MEM	:=TRUE;

	END_IF;
	IF LASER_SENSOR_2_IR THEN
		LASER_SENSOR_2_IR_MEM	:=TRUE;

	END_IF;
// PALLET STATION
	ACTUAL_PALLET_LIFTER_POS := ComTCP_SimInputs.pallet_lifter_AXIS;
	PALLET_FORK_ENABLED			:= ComTCP_SimInputs.pallet_fork_left_FB;
	PALLET_LIGHT_BARRIER_1		:= ComTCP_SimInputs.pallet_light_barrier_1_IR;
	PALLET_LIGHT_BARRIER_2		:= ComTCP_SimInputs.pallet_light_barrier_2_IR;
END_PROGRAM

PROGRAM _EXIT
	(* Insert code here *)

END_PROGRAM
```

#### Variables.var - Local variables
```iecst
VAR
	count3 : INT;
	count2 : INT;
	count : INT;
END_VAR
```

### Program Logical/Feeder_Handler (IEC)

#### Main.st - Init, cyclic, exit code
```iecst
PROGRAM _INIT
	(* Insert code here *)
	Carriage_2_target_position_array[0]:=0.44;
	Carriage_2_target_position_array[1]:=1.1;
	Carriage_2_target_position_array[2]:=0.9;
	index:=0;
	CountPusherState	:= 8;

END_PROGRAM

PROGRAM _CYCLIC
	(* Insert code here *)

	CASE State_Feeder OF
		WaitPowerON:
			IF POWER_ON_FEEDER THEN
			conveyor_if_disable_request	:= TRUE;
			conveyor_turn1_disable_request	:= TRUE;
			conveyor_end_disable_request	:= TRUE;
			carriage_2.PowerON				:=TRUE;
			State_Feeder							:=WaitStart;
			END_IF;

		WaitStart:
			IF (START_FEEDER) THEN
				conveyor_if_enable_request	:=TRUE;
				conveyor_end_enable_request	:=TRUE;
				conveyor_turn1_enable_request	:=TRUE;
				IF carriage_2.Powered THEN
					START_FEEDER				:= FALSE;
					POWER_ON_FEEDER 			:= FALSE;
					State_Feeder						:= WaitConveyorEnabled;
				END_IF;
			END_IF;
		WaitConveyorEnabled:

			IF NOT conveyor_if_enable_request AND NOT conveyor_end_enable_request AND NOT conveyor_turn1_enable_request THEN

				State_Feeder	:= WaitSensorBox;
			END_IF;

		WaitSensorBox:

			IF LASER_SENSOR_IR  THEN
//				LASER_SENSOR_IR_MEM	:= FALSE;
				COUNT_LASER_SENSOR_IR:=COUNT_LASER_SENSOR_IR+1;
				State_Feeder	:= WaitpusherenableStop;
			END_IF;

		WaitpusherenableStop:

			IF NOT WaitCarriage AND NOT FIRST_LAYER_OPERATION THEN

				IF NUM_BOX_COUNTED<=7 THEN
					pusher_enable_request	:= TRUE;
					State_Feeder	:= WaitPusherStop;
				END_IF;

				IF NUM_BOX_COUNTED=8 THEN
					pusher_enable_request	:= TRUE;
					FIRST_LAYER_OPERATION		:=TRUE;
					NUM_BOX_COUNTED :=0;
					State_Feeder	:= WaitPusherStop;
				END_IF;
  			END_IF;
			IF NOT WaitCarriage AND FIRST_LAYER_OPERATION THEN
				IF NUM_BOX_COUNTED<=5 THEN
					pusher_enable_request	:= TRUE;
					State_Feeder	:= WaitPusherStop;

				END_IF;

				IF NUM_BOX_COUNTED=6 THEN
					pusher_enable_request	:= TRUE;
					State_Feeder	:= WaitPusherStop;
				END_IF;
			END_IF;

		WaitPusherStop:
			IF ( NOT pusher_enable_request) THEN
				pusher_disable_request	:= TRUE;
				State_Feeder	:= WaitSensorCount;

			END_IF;

		WaitSensorCount:
			IF ( NOT pusher_disable_request)AND LASER_SENSOR_2_IR_MEM THEN
				LASER_SENSOR_2_IR_MEM	:= FALSE;
				ACTUAL_BOXES := ACTUAL_BOXES  + 1;
				NUM_BOX_COUNTED := NUM_BOX_COUNTED + 1;
				COUNT_BOXES_NUMBER	:= COUNT_BOXES_NUMBER+1;
				CountPusherState	:= CountPusherState + 1;
				IF NOT FIRST_LAYER_OPERATION THEN

					IF NUM_BOX_COUNTED=8  THEN
						WaitCarriage				:= TRUE;
						IF NOT oddsequence  THEN
	  						FIRST_LAYER_OPERATION	:= NOT FIRST_LAYER_OPERATION;
						END_IF;

						NUM_BOX_COUNTED :=0;
						TimeCount:=150;
						TimeOut								:= FALSE;
						State_Feeder	:=WaitCheckTurnPusher;
					ELSE
						conveyor_if_enable_request		:=TRUE;
						State_Feeder	:=  WaitConveyorEnabled;

					END_IF;

				ELSE
					IF NUM_BOX_COUNTED=3 OR NUM_BOX_COUNTED=6   THEN

						IF (oddsequence AND NUM_BOX_COUNTED=6) OR (oddsequence AND NUM_BOX_COUNTED>3) THEN

							FIRST_LAYER_OPERATION	:= NOT FIRST_LAYER_OPERATION;
							NUM_BOX_COUNTED :=0;
						END_IF;
						TimeCount		:=150;
						TimeOut			:= FALSE;
						WaitCarriage				:= TRUE;
						State_Feeder	:= WaitCheckTurnPusher;
					ELSE
						conveyor_if_enable_request		:=TRUE;
						State_Feeder	:= WaitConveyorEnabled;

					END_IF;
				END_IF;
			END_IF;

		WaitCheckTurnPusher:

			IF CountPusherState = 16  THEN
				turnpusher_enable_request	:= TRUE;
				CountPusherState 			:= 0;

			END_IF;
			IF CountPusherState = 12  THEN
				CountPusherState 			:= 0;
				turnpusher_disable_request	:= TRUE;
			END_IF;
			IF ACTUAL_BOXES<14 THEN
				index:=0;
			ELSE
				index:=1;
				FEERDER_WAIT_TO_DELIVER_BOXES :=TRUE;
			END_IF;

			State_Feeder	:= WaitConveyor_endStop;

		WaitConveyor_endStop:

			TimeCount := TimeCount-1;

			IF TimeOut AND NOT FEEDER_ON_PHASE_STOP_WAIT AND NOT FEERDER_WAIT_TO_DELIVER_BOXES THEN

				carriage_2.Input_Target_Position 	:=Carriage_2_target_position_array[index];
				carriage_2.Actual_Command 			:= TARGETPOSITION;
				TimeOut								:= FALSE;
				State_Feeder	:= WaitCarriage_position;
			END_IF;

		WaitCarriage_position:
			IF carriage_2.InPosition THEN
				carriage_2.Actual_Command := HOMING;
				State_Feeder	:= WaitCarriage_Homing;
			END_IF;

		WaitCarriage_Homing:
			IF ((carriage_2.InPosition)AND (ACTUAL_BOXES<14)) THEN
				WaitCarriage				:= FALSE;
				State_Feeder	:= WaitConveyorEnabled;
			END_IF;
			IF (carriage_2.InPosition AND (ACTUAL_BOXES=14)) THEN
				oddsequence:= NOT oddsequence;
				FEERDER_BOXES_DELIVERED :=TRUE;
				ACTUAL_BOXES:=0;
			END_IF;
			IF (NOT carriage_2.InVelocity AND START_AGAIN_FEEDER) THEN
				START_AGAIN_FEEDER		:= FALSE;
				NUM_BOX_COUNTED			:=	0;
				WaitCarriage			:= FALSE;
				State_Feeder			:= WaitConveyorEnabled;
			END_IF;

		WaitStopSequence:
			IF  NOT pusher_disable_request AND NOT conveyor_turn1_disable_request AND NOT conveyor_end_disable_request  AND NOT carriage_2.InVelocity  THEN
				pusher_disable_request			:= TRUE;
				turnpusher_disable_request		:= TRUE;
				FEEDER_EMERGENCY_STOP	:= FALSE;
				FEEDER_IMMEDIATE_STOP	:= FALSE;
				FEEDER_ON_PHASE_STOP	:= FALSE;
				START_FEEDER			:= FALSE;

				IF emergency_stop  THEN
					emergency_stop := FALSE;
					FIRST_LAYER_OPERATION			:= FALSE;
					COUNT_BOXES_NUMBER				:=0;
					NUM_BOX_COUNTED					:= 0;
					ACTUAL_BOXES					:= 0;
	  				State_Feeder			:= WaitPowerON;
				ELSE
					State_Feeder			:= WaitStart;
				END_IF;

			END_IF;

			IF Stop_all THEN

				conveyor_if_disable_request		:= TRUE;
				conveyor_turn1_disable_request	:= TRUE;
				conveyor_end_disable_request	:= TRUE;
				carriage_2.Actual_Command 		:= POWEROFF;
				pusher_disable_request			:= TRUE;
				turnpusher_disable_request		:= TRUE;
				FIRST_LAYER_OPERATION			:= FALSE;
				COUNT_BOXES_NUMBER				:=0;
				NUM_BOX_COUNTED					:= 0;
				ACTUAL_BOXES					:= 0;
				Stop_all						:= TRUE;
				State_Feeder					:= WaitPowerON;
			END_IF;

	END_CASE
	IF FEEDER_STOP THEN
		FEEDER_STOP	:= FALSE;
		Stop_all	:= TRUE;
		State_Feeder					:= WaitStopSequence;
	END_IF;
	IF FEEDER_EMERGENCY_STOP OR FEEDER_IMMEDIATE_STOP THEN
		emergency_stop := TRUE;
		conveyor_if_disable_request		:= TRUE;
		conveyor_turn1_disable_request	:= TRUE;
		conveyor_end_disable_request	:= TRUE;
		carriage_2.Actual_Command 		:= STOP;

		State_Feeder					:= WaitStopSequence;
	END_IF;
	IF FEEDER_ON_PHASE_STOP THEN
		FEEDER_ON_PHASE_STOP_WAIT 	:= TRUE;
		FEEDER_ON_PHASE_STOP		:= FALSE;
	END_IF;

	IF  TimeCount = 0 THEN
		TimeOut := TRUE;

	END_IF;

	conveyor_if.DeviceOperation := OperationType;
	conveyor_if.DeviceClock := TRUE;
	conveyor_if.DeviceDiagnosticsEnabled := TRUE;
	conveyor_if.DeviceEnablePreset := FALSE;
	conveyor_if.DeviceEnableTime := 10;
	conveyor_if.DeviceDisableTime := 10;
	conveyor_if.DeviceType := DEVICE_WITHOUT_FEEDBACK OR DEVICE_WITH_SINGLE_ACTUATION;
	conveyor_if(DeviceEnableRequest := conveyor_if_enable_request, DeviceDisableRequest := conveyor_if_disable_request );
	ENABLE_CONVEYOR_IF:= conveyor_if.EnableDevice;
	// fault generation is directly manage in signal mnagement since it will desactivated
	CONVEYOR_IF_FAULT:= conveyor_if.DeviceFault;

	pusher.DeviceOperation := OperationType;
	pusher.DeviceClock := TRUE;
	pusher.DeviceDiagnosticsEnabled := TRUE;
	pusher.DeviceEnablePreset := FALSE;
	pusher.DeviceEnabledSensor := PUSHER_ENABLED;
	pusher.DeviceDisabledSensor := PUSHER_DISABLED;
	pusher.DeviceEnableTime := 10;
	pusher.DeviceDisableTime := 10;
	pusher.DeviceType := DEVICE_WITH_DOUBLE_FEEDBACK OR DEVICE_WITH_SINGLE_ACTUATION;
	pusher(DeviceEnableRequest := pusher_enable_request, DeviceDisableRequest := pusher_disable_request );
	ENABLE_PUSHER:= pusher.EnableDevice;
	pusher.SimulationDeviceFault := SIMULATE_FAULT_PUSHER;
	PUSHER_FAULT:= (pusher.DeviceFault AND POWER_MACHINE);

	turnpusher.DeviceOperation := OperationType;
	turnpusher.DeviceClock := TRUE;
	turnpusher.DeviceDiagnosticsEnabled := TRUE;
	turnpusher.DeviceEnablePreset := FALSE;
	turnpusher.DeviceEnabledSensor := TURNPUSHER_ENABLED;
	turnpusher.DeviceDisabledSensor := TURNPUSHER_DISABLED;
	turnpusher.DeviceEnableTime := 100;
	turnpusher.DeviceDisableTime := 100;
	turnpusher.DeviceType := DEVICE_WITH_DOUBLE_FEEDBACK OR DEVICE_WITH_DOUBLE_ACTUATION;
	turnpusher(DeviceEnableRequest := turnpusher_enable_request, DeviceDisableRequest := turnpusher_disable_request );
	ENABLE_TURNPUSHER:= turnpusher.EnableDevice;
	DISABLE_TURNPUSHER := turnpusher.DisableDevice;
	turnpusher.SimulationDeviceFault := SIMULATE_FAULT_TURNPUSHER;
	TURNPUSHER_FAULT := (turnpusher.DeviceFault AND POWER_MACHINE);

	conveyor_turn1.DeviceOperation := OperationType;
	conveyor_turn1.DeviceClock := TRUE;
	conveyor_turn1.DeviceDiagnosticsEnabled := TRUE;
	conveyor_turn1.DeviceEnablePreset := FALSE;
	conveyor_turn1.DeviceEnableTime := 100;
	conveyor_turn1.DeviceDisableTime := 50;
	conveyor_turn1.DeviceType := DEVICE_WITHOUT_FEEDBACK OR DEVICE_WITH_SINGLE_ACTUATION;
	conveyor_turn1(DeviceEnableRequest := conveyor_turn1_enable_request, DeviceDisableRequest := conveyor_turn1_disable_request );
	ENABLE_CONVEYOR_TURN1 := conveyor_turn1.EnableDevice;

	// fault generation is directly manage in signal mnagement since it will desactivated
	CONVEYOR_TURN1_FAULT := conveyor_turn1.DeviceFault;

	conveyor_end.DeviceOperation := OperationType;
	conveyor_end.DeviceClock := TRUE;
	conveyor_end.DeviceDiagnosticsEnabled := TRUE;
	conveyor_end.DeviceEnablePreset := FALSE;
	conveyor_end.DeviceEnableTime := 100;
	conveyor_end.DeviceDisableTime := 50;
	conveyor_end.DeviceType := DEVICE_WITHOUT_FEEDBACK OR DEVICE_WITH_SINGLE_ACTUATION;
	conveyor_end(DeviceEnableRequest := conveyor_end_enable_request, DeviceDisableRequest := conveyor_end_disable_request );
	ENABLE_CONVEYOR_END := conveyor_end.EnableDevice;

	// fault generation is directly manage in signal mnagement since it will desactivated
	CONVEYOR_END_FAULT := conveyor_end.DeviceFault;

	carriage_2.DeviceClock := TRUE;
	carriage_2.DeviceTimer := 100;
	carriage_2.Reached_Postion:= CARRIAGE_RCHD_POS;
	carriage_2.DeviceFeedback := TRUE;
	carriage_2.InputSimulateError:=SIMULATE_FAULT_CARRIAGE_2; //input of fault then name
	CARRIAGE_2_FAULT:= carriage_2.OutputSimulateError;
	carriage_2.Actual_position:= ACTUAL_CARRIAGE_POS;
	CARRIAGE_TRG_POS := carriage_2.Output_Target_Position;
	carriage_2();

END_PROGRAM

PROGRAM _EXIT
	(* Insert code here *)

END_PROGRAM
```

#### Types.typ - Local data types
```iecst
TYPE
	FeederStateType :
	(
		WaitPowerON,
		WaitStart,
		WaitConveyorEnabled,
		WaitSensorBox,
		WaitpusherenableStop,
		WaitPusherStop,
		WaitSensorCount,
		WaitConveyor_endStop,
		WaitCheckTurnPusher,
		WaitCarriage_position,
		WaitCarriage_Homing,
		WaitStopSequence

	);
END_TYPE
```

#### Variables.var - Local variables
```iecst
VAR
	conveyor_if : Generic_Device;
	conveyor_end : Generic_Device;
	conveyor_end_enable_request : BOOL;
	conveyor_end_disable_request : BOOL;
	conveyor_turn1 : Generic_Device;
	conveyor_turn1_enable_request : BOOL;
	conveyor_turn1_disable_request : BOOL;
	turnpusher : Generic_Device;
	turnpusher_enable_request : BOOL;
	turnpusher_disable_request : BOOL;
	pusher : Generic_Device;
	pusher_enable_request : BOOL;
	pusher_disable_request : BOOL;
	conveyor_if_enable_request : BOOL;
	conveyor_if_disable_request : BOOL;
	State_Feeder : FeederStateType;
	Carriage_2_target_position_array : ARRAY[0..2] OF REAL;
	carriage_2 : Generic_Axis;
	carriage_actual_command : DWORD;
	index : INT;
	carriageTiming : INT := 10;
	oddsequence : BOOL; (*used to invert the next sequence of boxes*)
	emergency_stop : BOOL;
	TimeOut : BOOL;
	TimeCount : INT;
	WaitCarriage : BOOL;
	CountPusherState : INT;
	TURNPUSHER_DISABLED_1111 : BOOL;
	Stop_all : BOOL;
END_VAR
```

### Program Logical/Crane_Handler (IEC)

#### Main.st - Init, cyclic, exit code
```iecst
PROGRAM _INIT
	(* Insert code here *)
	gantrycranetarget_position_array[0]:= -1.11;
	gantrycranetarget_position_array[1]:= -1.3;
	index_gantry_crane:=0;

	box_crane_target_position_array[0]:= 0.01;
	box_crane_target_position_array[1]:= -0.195;
	box_crane_target_position_array[2]:= -0.2;
	index_box_crane:=0;

END_PROGRAM

PROGRAM _CYCLIC
	(* Insert code here *)
	CASE State_Crane OF

		WaitPowerON:
			IF POWER_ON_CRANE THEN

				slide_rail_right_disable_request	:= TRUE;
				vacuum_box_crane_disable_request	:= TRUE;
				pusher_x_disable_request			:= TRUE;
				pusher_z_disable_request			:= TRUE;
				cartborad_disable_request			:= TRUE;
				box_crane.PowerON					:= TRUE;
				gantry_crane.PowerON				:= TRUE;
				State_Crane							:=WaitStart;
			END_IF;
		WaitStart:
			IF (START_CRANE AND NOT StartAgain) THEN
				START_CRANE		:= FALSE;
				State_Crane		:= WaitBox_craneMove;
			END_IF;
			IF (START_CRANE AND StartAgain) THEN
				StartAgain		:= FALSE;
	  			State_Crane		:= Crane_immediate_stop;
			END_IF;

		WaitBox_craneMove:
			IF NOT first_layer_release_CB AND NOT gantry_crane.InVelocity THEN
				Crane_immediate_stop := 2;
				index_box_crane					:= 1;
				IF box_crane.Powered THEN
					box_crane.Input_Target_Position := box_crane_target_position_array[index_box_crane];
					box_crane.Actual_Command		:= TARGETPOSITION;
					State_Crane						:= WaitTakeReleaseCartboard;
				END_IF;
			END_IF;

			IF first_layer_release_CB AND NOT box_crane.InVelocity AND NOT gantry_crane.InVelocity THEN
				Crane_immediate_stop := 6;
				index_box_crane					:= 2;
				first_layer_release_CB			:= FALSE;
				box_crane.Input_Target_Position := box_crane_target_position_array[index_box_crane];
				box_crane.Actual_Command		:= TARGETPOSITION;
				release_cartboard				:= TRUE;
				State_Crane						:= WaitTakeReleaseCartboard;

			END_IF;

		WaitBox_craneMoveNEW:

			IF second_layer_release_CB  THEN
				Crane_immediate_stop := 6;
				IF  NOT pusher_z_enable_request AND NOT slide_rail_right_enable_request  THEN
					index_box_crane					:= 0;
					second_layer_release_CB			:= FALSE;
					box_crane.Input_Target_Position := box_crane_target_position_array[index_box_crane];
					box_crane.Actual_Command		:= TARGETPOSITION;
					box_crane_upper_position		:= TRUE;
					State_Crane						:= WaitBox_craneMoveNEW;
				END_IF;
			END_IF;
			IF box_crane_upper_position	AND  box_crane.InPosition THEN
				Crane_immediate_stop := 6;
				box_crane_upper_position		:= FALSE;
				release_cartboard				:= TRUE;
				Box_craneMoveNEW				:= TRUE;
				State_Crane						:= WaitGantry_craneMove;
			END_IF;
		WaitTakeReleaseCartboard:

			IF (NOT release_cartboard AND NOT CRANE_ON_PHASE_STOP_WAIT ) THEN
				Crane_immediate_stop := 4;
				IF box_crane.InPosition THEN
					cartborad_enable_request			:= TRUE;
					vacuum_box_crane_enable_request		:= TRUE;
					State_Crane						:= WaitBox_craneTakeHome;
				END_IF;
			END_IF;

			IF (release_cartboard AND gantry_crane.InPosition ) OR (release_cartboard AND NOT box_crane.InVelocity AND NOT Box_craneMoveNEW ) THEN
				Crane_immediate_stop := 6;
				release_cartboard					:= FALSE;
				Box_craneMoveNEW					:= FALSE;
				vacuum_box_crane_disable_request	:= TRUE;
				cartborad_disable_request			:= TRUE;
				release_boxes						:= TRUE;
				State_Crane							:= WaitGantry_craneMove;
			END_IF;

		WaitBox_craneTakeHome:
			Crane_immediate_stop := 4;
			IF NOT cartborad_enable_request AND NOT vacuum_box_crane_enable_request THEN
				box_crane.Actual_Command		:= HOMING;
				CRANE_WAIT_BOXES				:= TRUE;
				COUNT_CARTBOARD_NUMBER				:= COUNT_CARTBOARD_NUMBER-1;
				SECOND_LAYER_OPERATION			:= NOT SECOND_LAYER_OPERATION;
				State_Crane						:= WaitBox_craneBoxes;
			END_IF;
		WaitBox_craneBoxes:
			Crane_immediate_stop := 5;
			IF NOT box_crane.InVelocity AND NOT CRANE_WAIT_BOXES  THEN
				pusher_z_enable_request			:= TRUE;
				slide_rail_right_enable_request	:= TRUE;
				IF NOT SECOND_LAYER_OPERATION THEN
					second_layer_release_CB			:= TRUE;
					State_Crane						:= WaitBox_craneMoveNEW;

				ELSE
					State_Crane						:= WaitGantry_craneMove;
				END_IF;

			END_IF;

		WaitGantry_craneMove:

			IF NOT release_boxes AND NOT cartborad_enable_request AND NOT vacuum_box_crane_enable_request THEN
				Crane_immediate_stop := 6;
				IF NOT pusher_z_enable_request AND NOT slide_rail_right_enable_request THEN
					index_gantry_crane := 0;
					gantry_crane.Input_Target_Position := gantrycranetarget_position_array[index_gantry_crane];
					gantry_crane.Actual_Command		:= TARGETPOSITION;

					IF NOT SECOND_LAYER_OPERATION OR Box_craneMoveNEW THEN
						(*Box_craneMoveNEW				:= FALSE;*)
						release_cartboard				:= TRUE;
						//nwe step
						State_Crane						:= WaitTakeReleaseCartboard;
					ELSE
						first_layer_release_CB			:= TRUE;
						State_Crane						:= WaitBox_craneMove;
					END_IF;

				END_IF;
			END_IF;

			IF release_boxes AND NOT cartborad_enable_request AND NOT vacuum_box_crane_enable_request THEN
				Crane_immediate_stop := 3;
				release_boxes						:= FALSE;
				index_gantry_crane 					:= 1;
				gantry_crane.Input_Target_Position  := gantrycranetarget_position_array[index_gantry_crane];
				gantry_crane.Actual_Command			:= TARGETPOSITION;
				State_Crane							:= WaitSlide_rail_rightMove;
			END_IF;

		WaitSlide_rail_rightMove:
			Crane_immediate_stop := 5;
			IF gantry_crane.InPosition THEN
				slide_rail_right_disable_request	:= TRUE;
				State_Crane							:= WaitGantry_cranePusher_xMove;
			END_IF;

		WaitGantry_cranePusher_xMove:
			Crane_immediate_stop := 9;
			IF  NOT slide_rail_right_disable_request THEN
	  			pusher_x_enable_request			:= TRUE;
				gantry_crane.Actual_Command		:= HOMING;

			State_Crane							:= WaitPusher_xPusher_zMove;
			END_IF;
		WaitPusher_xPusher_zMove:
			Crane_immediate_stop := 8;
			IF NOT gantry_crane.InVelocity AND NOT pusher_x_enable_request THEN
				pusher_x_disable_request		:= TRUE;
				pusher_z_disable_request		:= TRUE;
				CRANE_BOXES_DELIVERED			:= TRUE;
				State_Crane							:= WaitBox_craneMove;
			END_IF;

		WaitStopSequence:
			IF 	(NOT box_crane.InVelocity AND NOT gantry_crane.InVelocity)  THEN

				State_Crane					:= WaitStart;
			END_IF;

		WaitEmergenceStopSequence:
	END_CASE;

	IF CRANE_STOP THEN
		CRANE_STOP	:= FALSE;
		gantry_crane.Actual_Command 		:= POWEROFF;
		box_crane.Actual_Command 			:= POWEROFF;
		pusher_x_disable_request			:= TRUE;
		pusher_z_disable_request			:= TRUE;
		slide_rail_right_disable_request	:= TRUE;
		State_Crane							:= WaitPowerON;
	END_IF;

	IF CRANE_EMERGENCY_STOP THEN
		gantry_crane.Actual_Command 		:= STOP;
		box_crane.Actual_Command 			:= STOP;
		CRANE_EMERGENCY_STOP				:= FALSE;
		State_Crane							:= WaitStopSequence;
	END_IF;

	IF  CRANE_IMMEDIATE_STOP THEN
		StartAgain					:= TRUE;
		gantry_crane.Actual_Command 		:= STOP;
		box_crane.Actual_Command 			:= STOP;
		IF release_boxes THEN

		ELSIF ((SECOND_LAYER_OPERATION OR Box_craneMoveNEW) AND NOT release_boxes)   THEN

			IF NOT release_boxes  THEN
				SECOND_LAYER_OPERATION :=TRUE;
				Box_craneMoveNEW		:=TRUE;
			END_IF;
			State_Crane					:= WaitGantry_craneMove;
		ELSE
			State_Crane					:= WaitStart;
		END_IF;

	END_IF;
	IF CRANE_ON_PHASE_STOP THEN
		CRANE_ON_PHASE_STOP			:= FALSE;
		CRANE_ON_PHASE_STOP_WAIT 	:= TRUE;

	END_IF;

	slide_rail_right.DeviceOperation := OperationType;
	slide_rail_right.DeviceClock := TRUE;
	slide_rail_right.DeviceDiagnosticsEnabled := TRUE;
	slide_rail_right.DeviceEnablePreset := FALSE;
	slide_rail_right.DeviceEnableTime := 100;
	slide_rail_right.DeviceDisableTime := 100;
	slide_rail_right.DeviceType := DEVICE_WITHOUT_FEEDBACK OR DEVICE_WITH_SINGLE_ACTUATION;
	slide_rail_right(DeviceEnableRequest := slide_rail_right_enable_request, DeviceDisableRequest := slide_rail_right_disable_request );
	ENABLE_SLIDE_RAIL_RIGHT := slide_rail_right.EnableDevice;
	slide_rail_right.SimulationDeviceFault	:= SIMULATE_FAULT_SLIDE_RAIL_RIGHT;
	SLIDE_RAIL_RIGHT_FAULT := (slide_rail_right.DeviceFault AND POWER_MACHINE);

	vacuum_box_crane.DeviceOperation := OperationType;
	vacuum_box_crane.DeviceClock := TRUE;
	vacuum_box_crane.DeviceDiagnosticsEnabled := FALSE;
	vacuum_box_crane.DeviceEnablePreset := FALSE;
	vacuum_box_crane.DeviceEnabledSensor := VACUUM_BOX_CRANE_ENABLED;
	vacuum_box_crane.DeviceEnableTime := 20;
	vacuum_box_crane.DeviceDisableTime := 20;
	vacuum_box_crane.DeviceType := DEVICE_WITH_ENABLE_FEEDBACK OR DEVICE_WITH_SINGLE_ACTUATION;
	vacuum_box_crane(DeviceEnableRequest := vacuum_box_crane_enable_request, DeviceDisableRequest := vacuum_box_crane_disable_request );
	ENABLE_VACUUM_BOX_CRANE := vacuum_box_crane.EnableDevice;
	vacuum_box_crane.SimulationDeviceFault	:= SIMULATE_FAULT_VACUUM_BOX_CRANE;
	VACUUM_BOX_CRANE_FAULT := (vacuum_box_crane.DeviceFault AND POWER_MACHINE);

	pusher_x.DeviceOperation := OperationType;
	pusher_x.DeviceClock := TRUE;
	pusher_x.DeviceDiagnosticsEnabled := FALSE;
	pusher_x.DeviceEnablePreset := FALSE;
	pusher_x.DeviceEnableTime := 100;
	pusher_x.DeviceDisableTime := 100;
	pusher_x.DeviceType := DEVICE_WITHOUT_FEEDBACK OR DEVICE_WITH_SINGLE_ACTUATION;
	pusher_x(DeviceEnableRequest := pusher_x_enable_request, DeviceDisableRequest := pusher_x_disable_request );
	ENABLE_PUSHER_X := pusher_x.EnableDevice;
	pusher_x.SimulationDeviceFault	:= SIMULATE_FAULT_PUSHER_X;
	PUSHER_X_FAULT := ( pusher_x.DeviceFault AND POWER_MACHINE);

	pusher_z.DeviceOperation := OperationType;
	pusher_z.DeviceClock := TRUE;
	pusher_z.DeviceDiagnosticsEnabled := FALSE;
	pusher_z.DeviceEnablePreset := FALSE;
	pusher_z.DeviceEnableTime := 100;
	pusher_z.DeviceDisableTime := 100;
	pusher_z.DeviceType := DEVICE_WITHOUT_FEEDBACK OR DEVICE_WITH_SINGLE_ACTUATION;
	pusher_z(DeviceEnableRequest := pusher_z_enable_request, DeviceDisableRequest := pusher_z_disable_request );
	ENABLE_PUSHER_Z := pusher_z.EnableDevice;
	pusher_z.SimulationDeviceFault	:= SIMULATE_FAULT_PUSHER_Z;
	PUSHER_Z_FAULT := (pusher_z.DeviceFault AND POWER_MACHINE);

	cartborad.DeviceOperation := OperationType;
	cartborad.DeviceClock := TRUE;
	cartborad.DeviceDiagnosticsEnabled := FALSE;
	cartborad.DeviceEnablePreset := FALSE;
	cartborad.DeviceEnableTime := 25;
	cartborad.DeviceDisableTime := 25;
	cartborad.DeviceType := DEVICE_WITHOUT_FEEDBACK OR DEVICE_WITH_SINGLE_ACTUATION;
	cartborad(DeviceEnableRequest := cartborad_enable_request, DeviceDisableRequest := cartborad_disable_request );
	ENABLE_CARTBORAD := cartborad.EnableDevice;
	cartborad.SimulationDeviceFault	:= SIMULATE_FAULT_CARTBORAD;
	CARTBORAD_FAULT := (cartborad.DeviceFault AND POWER_MACHINE);
	IF cartborad.DeviceFault THEN
		coutn := coutn + 1;

	END_IF;

	gantry_crane.DeviceClock := TRUE;
	gantry_crane.DeviceTimer := 100 ;
	gantry_crane.Reached_Postion:= GANTRY_CRANE_RCHD_POS;// no available without feedback
	gantry_crane.DeviceFeedback := FALSE;
	gantry_crane.InputSimulateError:=SIMULATE_FAULT_GANTRY_CRANE;
	GANTRY_CRANE_FAULT := gantry_crane.OutputSimulateError;
	gantry_crane.Actual_position:= ACTUAL_GANTRY_CRANE_POS;
	GANTRY_CRANE_TRG_POS := gantry_crane.Output_Target_Position;

	gantry_crane();

	box_crane.DeviceClock := TRUE;
	box_crane.DeviceTimer := 100 ;
	box_crane.Reached_Postion:= BOX_CRANE_RCHD_POS;// no available without feedback
	box_crane.DeviceFeedback := FALSE;
	box_crane.InputSimulateError:=SIMULATE_FAULT_BOX_CRANE;
	BOX_CRANE_FAULT := box_crane.OutputSimulateError ;
	box_crane.Actual_position:= ACTUAL_BOX_CRANE_POS;
	BOX_CRANE_TRG_POS := box_crane.Output_Target_Position;
	box_crane();

END_PROGRAM

PROGRAM _EXIT
	(* Insert code here *)

END_PROGRAM
```

#### Types.typ - Local data types
```iecst
TYPE
	CraneStateType :
		(
		WaitPowerON,
		WaitStart,
		WaitBox_craneMove,
		WaitBox_craneMoveNEW,
		WaitTakeReleaseCartboard,
		WaitBox_craneTakeHome,
		WaitBox_craneBoxes,
		WaitGantry_craneMove,
		WaitGantry_cranePusher_xMove,
		WaitSlide_rail_rightMove,
		WaitPusher_xPusher_zMove,
		WaitStopSequence,
		WaitEmergenceStopSequence

	);

END_TYPE
```

#### Variables.var - Local variables
```iecst
VAR
	slide_rail_right : Generic_Device;
	slide_rail_right_enable_request : BOOL;
	slide_rail_right_disable_request : BOOL;
	vacuum_box_crane : Generic_Device;
	vacuum_box_crane_enable_request : BOOL;
	vacuum_box_crane_disable_request : BOOL;
	pusher_x : Generic_Device;
	pusher_x_enable_request : BOOL;
	pusher_x_disable_request : BOOL;
	pusher_z : Generic_Device;
	pusher_z_enable_request : BOOL;
	pusher_z_disable_request : BOOL;
	cartborad : Generic_Device;
	cartborad_enable_request : BOOL;
	cartborad_disable_request : BOOL;
	box_crane : Generic_Axis;
	gantry_crane : Generic_Axis;
	box_crane_target_position_array : ARRAY[0..2] OF REAL;
	gantrycranetarget_position_array : ARRAY[0..1] OF REAL;
	index_box_crane : INT;
	index_gantry_crane : INT;
	State_Crane : CraneStateType;
	first_layer_release_CB : BOOL;
	second_layer_release_CB : BOOL;
	release_cartboard : BOOL;
	release_boxes : BOOL;
	box_crane_upper_position : BOOL;
	Box_craneMoveNEW : BOOL;
	Crane_immediate_stop : INT;
	StartAgain : BOOL;
	coutn : INT;
END_VAR
```

### Program Logical/Pallet_Handler (IEC)

#### Main.st - Init, cyclic, exit code
```iecst
PROGRAM _INIT
	(* Insert code here *)
	palletliftertargetposition_array[0]:= -0.12;
	palletliftertargetposition_array[1]:= -0.258;
	index_palletlifter:=0;

	pallet_convtarget_velocity_array[0]:= 0.1;
	pallet_convtarget_velocity_array[1]:= 0.5;
	index_pallet_conv:=0;
END_PROGRAM

PROGRAM _CYCLIC
	(* Insert code here *)

	CASE State_Pallet OF
		WaitPPowerON:
			IF POWER_ON_PALLET THEN

				pallet_conv_1_disable_request	:= TRUE;
				pallet_fork_disable_request 	:= TRUE;
				pallet_lifter.PowerON			:= TRUE;
				pallet_conveyor_2.PowerON		:= TRUE;
				State_Pallet							:=WaitPStart;
			END_IF;

		WaitPStart:
			IF (START_PALLET) THEN
				START_PALLET		:= FALSE;
				POWER_ON_PALLET		:= FALSE;
				State_Pallet		:= Waitpallet_lifterMove;
			END_IF;
			IF (START_PALLET AND AFTER_IMMEDIATE_STOP) THEN
				State_Pallet		:= pallet_immadiate_stop;
			END_IF;

		Waitpallet_lifterMove:
			pallet_immadiate_stop :=2;
			IF (pallet_lifter.Powered AND NOT odditeration )  THEN

				index_palletlifter	:=	1;
				pallet_lifter.Input_Target_Position	:= palletliftertargetposition_array[index_palletlifter];
				pallet_lifter.Actual_Command := TARGETPOSITION;
				State_Pallet		:= Waitpallet_forkMove;
			END_IF;

			IF (NOT pallet_fork_enable_request AND odditeration) OR (AFTER_IMMEDIATE_STOP AND odditeration) THEN
				index_palletlifter	:=	0;
				pallet_lifter.Input_Target_Position	:= palletliftertargetposition_array[index_palletlifter];
				pallet_lifter.Actual_Command := TARGETPOSITION;
				State_Pallet		:= Waitpallet_forkMove;
			END_IF;
		Waitpallet_forkMove:
			pallet_immadiate_stop 	:= 3;

			IF (pallet_lifter.InPosition AND NOT odditeration) OR (AFTER_IMMEDIATE_STOP AND  NOT odditeration)THEN
				pallet_fork_enable_request	:= TRUE;
				pallet_immadiate_stop 	:= 2;
				odditeration			:= NOT odditeration;
				State_Pallet			:= Waitpallet_lifterMove;
			END_IF;
			IF  (pallet_lifter.InPosition AND odditeration AND index_palletlifter = 0 ) OR (AFTER_IMMEDIATE_STOP AND odditeration)THEN

				pallet_fork_disable_request	:= TRUE;
				odditeration			:= NOT odditeration;
				pallet_immadiate_stop 	:= 4;
				State_Pallet			:= WaitpalletHome;
			END_IF;

		WaitpalletHome:
			pallet_immadiate_stop 	:= 4;
			IF NOT pallet_fork_disable_request	 OR (AFTER_IMMEDIATE_STOP) THEN
				pallet_lifter.Actual_Command := HOMING;
				TimerCount		:=50;
				Timedelay		:= FALSE;
				State_Pallet			:= Waitpallet_conveyor_1Move;
			END_IF;

		Waitpallet_conveyor_1Move:
			pallet_immadiate_stop 	:= 5;
			TimerCount := TimerCount-1;
			IF Timedelay OR (AFTER_IMMEDIATE_STOP) THEN
				index_pallet_conv						:= 1;
				pallet_conveyor_2.Input_Target_Velocity	:= pallet_convtarget_velocity_array[index_pallet_conv];
				pallet_conveyor_2.Actual_Command		:= TARGETVELOCITY;
				IF Takeoff_pallet  THEN
					Takeoff_pallet			:= FALSE;
	  				State_Pallet			:= Waitpallet_lifterMove;
				ELSE
					pallet_conv_1_enable_request	:= TRUE;
					State_Pallet			:= Waitlight_barrier_2;
				END_IF;

			END_IF;

		Waitlight_barrier_2:
			pallet_immadiate_stop 	:= 8;

			IF PALLET_LIGHT_BARRIER_2 AND pallet_conveyor_2.InVelocity AND NOT pallet_conv_1_enable_request THEN
				pallet_conv_1_disable_request := TRUE;
				index_pallet_conv		:= 0;
				pallet_immadiate_stop 	:= 7;
				pallet_conveyor_2.Input_Target_Velocity		:= pallet_convtarget_velocity_array[index_pallet_conv];
				pallet_conveyor_2.Actual_Command		:= TARGETVELOCITY;
				State_Pallet					:= Waitlight_barrier_1;
			END_IF;

		Waitlight_barrier_1:
			pallet_immadiate_stop 	:= 7;
			IF (PALLET_LIGHT_BARRIER_1 AND pallet_conveyor_2.InVelocity ) OR (AFTER_IMMEDIATE_STOP)  THEN
				COUNT_PALLET_NUMBER					:= COUNT_PALLET_NUMBER	-1;
				PALLET_WAIT_BOXES					:= TRUE;
				pallet_conveyor_2.Actual_Command	:= HOMING;
				State_Pallet						:= Waitcraneandstart;
			END_IF;

		Waitcraneandstart:
			pallet_immadiate_stop 		:= 9;
			IF (NOT pallet_conveyor_2.InVelocity AND NOT PALLET_WAIT_BOXES AND NOT PALLET_ON_PHASE_STOP_WAIT AND NOT pallet_conv_1_disable_request)  OR (AFTER_IMMEDIATE_STOP) OR (PHASE_STOP_WAIT)THEN
				Takeoff_pallet			:= TRUE;
				Timedelay				:= TRUE;
				PHASE_STOP_WAIT			:= FALSE;
				State_Pallet			:=  Waitpallet_conveyor_1Move;
			END_IF;

		WaitOnPhaseStopSequence:

			IF PALLET_ON_PHASE_STOP_REMOVE THEN	//special activation of motore 2 to remove the current pallet
				index_pallet_conv		:= 1;
				pallet_conveyor_2.Input_Target_Velocity		:= pallet_convtarget_velocity_array[index_pallet_conv];
				pallet_conveyor_2.Actual_Command		:= TARGETVELOCITY;
				IF NOT PALLET_ON_PHASE_STOP_WAIT THEN
					PHASE_STOP_WAIT					:= TRUE;
//					PALLET_WAIT_BOXES					:= FALSE;
					PALLET_ON_PHASE_STOP_REMOVE		:= FALSE;

					State_Pallet					:= Waitcraneandstart;
				END_IF;
			END_IF;
			IF PALLET_ON_PHASE_STOP_IDLE THEN
				PALLET_ON_PHASE_STOP_IDLE 		:= FALSE;
	  			State_Pallet					:= Waitcraneandstart;
			END_IF;

	END_CASE;
	IF  TimerCount = 0 THEN
		Timedelay := TRUE;
	END_IF;
	IF PALLET_STOP THEN
		PALLET_STOP	:= TRUE;
		pallet_lifter.Actual_Command			:= POWEROFF;
		pallet_conveyor_2.Actual_Command 		:= POWEROFF;
		pallet_conv_1_disable_request			:= TRUE;
		pallet_fork_disable_request				:= TRUE;
		State_Pallet							:= WaitPPowerON;
	END_IF;
	IF PALLET_EMERGENCY_STOP THEN
		pallet_lifter.Actual_Command			:= STOP;
		pallet_conveyor_2.Actual_Command 		:= STOP;
		pallet_conv_1_disable_request			:= TRUE;
		PALLET_EMERGENCY_STOP					:= FALSE;
		State_Pallet								:=WaitPPowerON;
	END_IF;

	IF  PALLET_IMMEDIATE_STOP THEN

		pallet_lifter.Actual_Command			:= STOP;
		pallet_conveyor_2.Actual_Command 		:= STOP;
		pallet_conv_1_disable_request	:= TRUE;
		AFTER_IMMEDIATE_STOP					:= TRUE;
		State_Pallet							:=WaitPPowerON;

	END_IF;
	IF PALLET_ON_PHASE_STOP THEN

		PALLET_ON_PHASE_STOP_WAIT 	:= TRUE;
		IF PALLET_WAIT_BOXES THEN
			PALLET_ON_PHASE_STOP				:= FALSE;
	  		State_Pallet					:= WaitOnPhaseStopSequence;
		END_IF;

	END_IF;

	pallet_conveyor_1.DeviceOperation := OperationType;
	pallet_conveyor_1.DeviceClock := TRUE;
	pallet_conveyor_1.DeviceDiagnosticsEnabled := TRUE;
	pallet_conveyor_1.DeviceEnablePreset := FALSE;
	pallet_conveyor_1.DeviceEnableTime := 25;
	pallet_conveyor_1.DeviceDisableTime := 25;
	pallet_conveyor_1.DeviceType := DEVICE_WITHOUT_FEEDBACK OR DEVICE_WITH_SINGLE_ACTUATION;
	pallet_conveyor_1(DeviceEnableRequest := pallet_conv_1_enable_request, DeviceDisableRequest := pallet_conv_1_disable_request );
	ENABLE_PALLET_CONVEYOR_1 := pallet_conveyor_1.EnableDevice;
	// fault generation is directly manage in signal mnagement since it will desactivated

	PALLET_CONVEYOR_1_FAULT := pallet_conveyor_1.SimulationDeviceFault;
	IF PALLET_CONVEYOR_1_FAULT THEN
		coutn := coutn + 1;

	END_IF;

	pallet_fork.DeviceOperation := OperationType;
	pallet_fork.DeviceClock := TRUE;
	pallet_fork.DeviceDiagnosticsEnabled := TRUE;
	pallet_fork.DeviceEnablePreset := FALSE;
	pallet_fork.DeviceEnabledSensor := PALLET_FORK_ENABLED;
	pallet_fork.DeviceEnableTime := 100;
	pallet_fork.DeviceDisableTime := 100;
	pallet_fork.DeviceType := DEVICE_WITH_ENABLE_FEEDBACK OR DEVICE_WITH_SINGLE_ACTUATION;
	pallet_fork(DeviceEnableRequest := pallet_fork_enable_request, DeviceDisableRequest := pallet_fork_disable_request );
	ENABLE_PALLET_FORK := pallet_fork.EnableDevice;
	pallet_fork.SimulationDeviceFault	:= SIMULATE_FAULT_PALLET_FORK;
	PALLET_FORK_FAULT := pallet_fork.SimulationDeviceFault (*pallet_fork.DeviceFault*);

	pallet_conveyor_2.DeviceClock := TRUE;
	pallet_conveyor_2.DeviceTimer := 10 ;
	pallet_conveyor_2.DeviceFeedback := FALSE;
	pallet_conveyor_2.InputSimulateError:=SIMULATE_FAULT_PALLET_CONVEYOR_2;
	PALLET_CONVEYOR_2_FAULT := pallet_conveyor_2.OutputSimulateError;
	PALLET_CONVEYOR_2_TRG_VEL := pallet_conveyor_2.Output_Target_Velocity;
	pallet_conveyor_2();

	pallet_lifter.DeviceClock := TRUE;
	pallet_lifter.DeviceTimer := 10 ;
	pallet_lifter.Reached_Postion:= PALLET_LIFTER_RCHD_POS; // no available without feedback
	pallet_lifter.DeviceFeedback := FALSE;
	pallet_lifter.InputSimulateError:=SIMULATE_FAULT_PALLET_LIFTER;
	PALLET_LIFTER_FAULT := pallet_lifter.OutputSimulateError;
	pallet_lifter.Actual_position:= ACTUAL_PALLET_LIFTER_POS;
	PALLET_LIFTER_TRG_POS := pallet_lifter.Output_Target_Position;
	pallet_lifter();

END_PROGRAM

PROGRAM _EXIT
	(* Insert code here *)

END_PROGRAM
```

#### Types.typ - Local data types
```iecst
TYPE

	palletStateType :
		(
		WaitPPowerON,
		WaitPStart,
		Waitpallet_lifterMove,
		Waitpallet_forkMove,
		WaitpalletHome,
		Waitpallet_conveyor_1Move,
		Waitpallet_conveyor_2Move,
		Waitlight_barrier_1,
		Waitlight_barrier_2,
		Waitcraneandstart,
		WaitOnPhaseStopSequence,
		WaitEmergenceStopSequence

	);
END_TYPE
```

#### Variables.var - Local variables
```iecst
VAR
	pallet_lifter : Generic_Axis;
	pallet_conveyor_2 : Generic_Axis;
	pallet_fork : Generic_Device;
	pallet_fork_enable_request : BOOL;
	pallet_fork_disable_request : BOOL;
	pallet_conveyor_1 : Generic_Device;
	pallet_conv_1_enable_request : BOOL;
	pallet_conv_1_disable_request : BOOL;
	index_pallet_conv : INT;
	pallet_convtarget_velocity_array : ARRAY[0..1] OF REAL;
	index_palletlifter : INT;
	palletliftertargetposition_array : ARRAY[0..1] OF REAL;
	State_Pallet : palletStateType;
	odditeration : BOOL;
	Takeoff_pallet : BOOL;
	Timedelay : BOOL;
	TimerCount : INT;
	pallet_immadiate_stop : INT;
	coutn : INT;
	PHASE_STOP_WAIT : BOOL;
END_VAR
```

### Program Logical/MASTER (IEC)

#### Main.st - Init, cyclic, exit code
```iecst
PROGRAM _INIT
	(* Insert code here *)

END_PROGRAM

PROGRAM _CYCLIC
	(* Insert code here *)

	CASE State_Master OF

		Initialization:

  			POWER_ON_FEEDER			:= TRUE;
			POWER_ON_CRANE			:= TRUE;
			POWER_ON_PALLET			:= TRUE;
			BUTTON_START			:= FALSE;
			blink_start				:= FALSE;

			BUTTON_STOP				:= FALSE;
			blink_stop				:= FALSE;

			BUTTON_EMERGENCY_STOP	:= FALSE;
			blink_ermergency		:= FALSE;

			BUTTON_IMMEDIATE_STOP	:= FALSE;
			blink_immediatestop		:= FALSE;

			BUTTON_ON_PHASE_STOP	:= FALSE;
			blink_onphasestop		:= FALSE;

			BUTTON_INITIALIZATION	:= FALSE;
			blink_Fauld				:= FALSE;

			State_Master			:= WaitButtonStart;

		WaitButtonStart:

			IF BUTTON_START THEN
				OperationType		:= 1;
				blink_start			:= TRUE;
				blink_stop			:= TRUE;
				PalletOnPhaseStop	:= FALSE;
				CardboardOnPhaseStop	:= FALSE;
				CRANE_ON_PHASE_STOP_WAIT := FALSE;
				PALLET_ON_PHASE_STOP_WAIT	:= FALSE;
				FEEDER_ON_PHASE_STOP_WAIT 	:= FALSE;
				IF NOT AfterOnPhase THEN
					START_FEEDER		:= TRUE;
					START_CRANE			:= TRUE;
					START_PALLET		:= TRUE;
					AfterOnPhase		:= FALSE;
				END_IF;
				State_Master		:= WaitCheckHandlersStart;
			END_IF;

		WaitCheckHandlersStart:

			IF NOT START_FEEDER AND NOT START_CRANE AND NOT START_PALLET  THEN

				State_Master		:= WaitFeederFeedback;
			END_IF;

		WaitFeederFeedback:

			IF FEERDER_WAIT_TO_DELIVER_BOXES THEN
				Onelayeroperation		:=1;
				State_Master			:= WaitCraneFeedback;
			END_IF;

		WaitCraneFeedback:
			IF  (CRANE_WAIT_BOXES AND Onelayeroperation = 1) THEN

				IF CardboardOnPhaseStop THEN
					FEEDER_ON_PHASE_STOP			:= TRUE;
					CRANE_ON_PHASE_STOP				:= TRUE;
					State_Master		:= WaitOnphaseStop;
				END_IF;

				State_Master			:= WaitPalletFeedback;

			END_IF;
		WaitPalletFeedback:
			IF PALLET_WAIT_BOXES THEN
				IF Onelayeroperation = 1 THEN
					Carriage_start_moving			:= TRUE;

					FEERDER_WAIT_TO_DELIVER_BOXES	:= FALSE;
					State_Master					:= WaitFeederFeedback2;
				END_IF;
			END_IF;

		WaitFeederFeedback2:
			IF FEERDER_BOXES_DELIVERED AND NOT START_AGAIN_FEEDER THEN
				Carriage_start_moving		:= TRUE;
				START_AGAIN_FEEDER		:=TRUE;
				FEERDER_BOXES_DELIVERED	:=FALSE;
				Onelayeroperation 		:= 2;
				State_Master			:= WaitCraneFeedback2;
			END_IF;

		WaitCraneFeedback2:
			IF  (CRANE_WAIT_BOXES AND Onelayeroperation = 2) THEN

				IF Onelayeroperation = 2 THEN
					CRANE_WAIT_BOXES	:= FALSE;//there are boxes go next
				END_IF;
				CRANE_WAIT_BOXES	:= FALSE;//moi new
				IF CardboardOnPhaseStop THEN
					FEEDER_ON_PHASE_STOP			:= TRUE;
					CRANE_ON_PHASE_STOP				:= TRUE;
					State_Master		:= WaitOnphaseStop;
				END_IF;
				State_Master			:= WaitPalletFeedback2;
			END_IF;

		WaitPalletFeedback2:
			IF PALLET_WAIT_BOXES THEN
				IF Onelayeroperation = 2 AND CRANE_BOXES_DELIVERED THEN

					TwolayerOperation				:= TwolayerOperation + 1;
					IF TwolayerOperation = 2 THEN
						PALLET_WAIT_BOXES				:= FALSE;
						TwolayerOperation				:= TwolayerOperation - 2;
					END_IF;
					CRANE_BOXES_DELIVERED			:= FALSE;
					Onelayeroperation 				:= 0;
					State_Master					:= WaitFeederFeedback;
				END_IF;

			END_IF;
		WaitOnphaseStop:

			IF  PALLET_WAIT_BOXES AND CardboardOnPhaseStop AND TwolayerOperation = 2 THEN
	  			CRANE_BOXES_DELIVERED			:= FALSE;
				PALLET_WAIT_BOXES				:= FALSE;
				PALLET_ON_PHASE_STOP_REMOVE		:= FALSE;
				State_Master			:= WaitButtonStart;
			END_IF;
			BUTTON_START 			:=FALSE;
			State_Master			:= WaitButtonStart;

		WaitStopSequence:
			BUTTON_STOP	:= FALSE;
			BUTTON_START :=FALSE;
			FEEDER_STOP	:= TRUE;
			CRANE_STOP	:= TRUE;
			PALLET_STOP	:= TRUE;
			State_Master			:= Initialization;

	END_CASE;

	IF BUTTON_STOP THEN
		FEEDER_IMMEDIATE_STOP	:= TRUE;
		CRANE_IMMEDIATE_STOP	:= TRUE;
		PALLET_IMMEDIATE_STOP	:= TRUE;

		State_Master			:= WaitStopSequence;
	END_IF;
	// DIRECT COMMAND OF STOP
	IF SM_EMERGENCY_STOP THEN
 		FEEDER_EMERGENCY_STOP	:= TRUE;
		CRANE_EMERGENCY_STOP	:= TRUE;
		PALLET_EMERGENCY_STOP	:= TRUE;
		BUTTON_START 			:=FALSE;
		State_Master			:= Initialization;
	END_IF;

	IF SM_IMMEDIATE_STOP THEN
		FEEDER_IMMEDIATE_STOP	:= TRUE;
		CRANE_IMMEDIATE_STOP	:= TRUE;
		PALLET_IMMEDIATE_STOP	:= TRUE;
		BUTTON_START 			:=FALSE;
		State_Master					:= WaitButtonStart;
	END_IF;

	IF SM_ON_PHASE_STOP THEN
		FEEDER_ON_PHASE_STOP			:= TRUE;
		CRANE_ON_PHASE_STOP				:= TRUE;
		PALLET_ON_PHASE_STOP			:= TRUE;
		PALLET_ON_PHASE_STOP_IDLE		:= TRUE;
		BUTTON_START 					:= FALSE;
		AfterOnPhase					:= TRUE;
		State_Master					:= WaitButtonStart;
	END_IF;

	IF SM_IMMEDIATE_STOP_CAT1 THEN
		FEEDER_IMMEDIATE_STOP	:= TRUE;
		IF FEERDER_WAIT_TO_DELIVER_BOXES THEN
			CRANE_IMMEDIATE_STOP	:= TRUE;
		ELSE
			CRANE_ON_PHASE_STOP				:= TRUE;
		END_IF;
		PALLET_ON_PHASE_STOP			:= TRUE;
		BUTTON_START 					:=FALSE;
		State_Master					:= WaitButtonStart;
	END_IF;

	IF SM_ON_PHASE_STOP_CAT1 THEN
		BUTTON_START 			:=FALSE;
		CardboardOnPhaseStop	:= TRUE;
	END_IF;

END_PROGRAM

PROGRAM _EXIT
	(* Insert code here *)

END_PROGRAM
```

#### Types.typ - Local data types
```iecst
TYPE
	MasterStateType :
		(
		Initialization,
		WaitButtonStart,
		WaitCheckHandlersStart,
		WaitFeederFeedback,
		WaitCraneFeedback,
		WaitPalletFeedback,
		WaitFeederFeedback2,
		WaitCraneFeedback2,
		WaitPalletFeedback2,
		WaitOnphaseStop,
		WaitImmediateStop,
		WaitEmergenceStop,
		WaitStopSequence,
		WaitReinitializationSequence

	);

END_TYPE
```

#### Variables.var - Local variables
```iecst
VAR
	State_Master : MasterStateType;
	Onelayeroperation : INT;
	TwolayerOperation : INT;
	Carriage_start_moving : BOOL;
	PalletOnPhaseStop : BOOL;
	CardboardOnPhaseStop : BOOL;
	AfterOnPhase : BOOL;
END_VAR
```

### Program Logical/SignalManagement (IEC)

#### Main.st - Init, cyclic, exit code
```iecst
PROGRAM _INIT
	(* Insert code here *)

END_PROGRAM

PROGRAM _CYCLIC
	(* Insert code here *)
									//######### INITIALIZATIONS #################//
	IF (OperationType = INIT) THEN
		SignalManagement (OperationType := INIT);
		SignalManagement (OperationType := START_CONFIGURATION);
		SignalManagement.OperationType := CONFIGURATION;
//		OperationType := RUN;
	ELSE
		SignalManagement (OperationType := START_GENERATION);
		SignalManagement.OperationType := GENERATION;

		IF COUNT_CARTBOARD_NUMBER = 1 THEN
			boxcrane_Cartboard_ALMOST_FINISH := TRUE;
		ELSE
			boxcrane_Cartboard_ALMOST_FINISH := FALSE;
		END_IF;
		SignalManagement
			(SignalType := WARNING,
			SignalCode := ID_Cartboard_ALMOST_FINISH,
		SignalOutput := NONE OR MATERIALS_RUN_OUT_LAMP OR NONE,
		ActivationSignal := boxcrane_Cartboard_ALMOST_FINISH);
		IF COUNT_CARTBOARD_NUMBER = 0 THEN
			boxcrane_Cartboard_FINISH := TRUE;
		END_IF;
		SignalManagement
			(SignalType := ALARM OR AUTO_CONDITIONED_RESET,
			SignalCode := ID_Cartboard_FINISH,
		SignalOutput := ON_PHASE_STOP OR NONE OR NONE,
		ActivationSignal := boxcrane_Cartboard_FINISH);

		//######### HANDLING SIGNAL OF PALLET #################//
		IF COUNT_PALLET_NUMBER = 1 THEN
			pallet_lifter_ALMOST_FINISH := TRUE;
		ELSE
			pallet_lifter_ALMOST_FINISH := FALSE;
		END_IF;
		SignalManagement
			(SignalType := WARNING,
			SignalCode := ID_P_lifter_ALMOST_FINISH,
		SignalOutput := NONE OR MATERIALS_RUN_OUT_LAMP OR NONE,
		ActivationSignal := pallet_lifter_ALMOST_FINISH);

		IF COUNT_PALLET_NUMBER =0 THEN
			pallet_lifter_FINISH := TRUE;
		END_IF;

		SignalManagement
			(SignalType := ALARM OR AUTO_CONDITIONED_RESET,
			SignalCode := ID_pallet_lifter_FINISH,
		SignalOutput := ON_PHASE_STOP OR NONE OR NONE,
		ActivationSignal := pallet_lifter_FINISH);

		//######### BUTTON HANDLING SIGNALS #################//
		//EMERGENCY STOP
		SignalManagement
			(SignalType := ALARM,
			SignalCode := ID_EMERGENCY_STOP,
		SignalOutput := EMERGENCY_STOP OR NONE OR NONE,
		ActivationSignal := BUTTON_EMERGENCY_STOP);

		//IMMEDIATE STOP
		SignalManagement
			(SignalType := ALARM,
			SignalCode := ID_IMMEDIATE_STOP,
		SignalOutput := IMMEDIATE_STOP OR NONE OR NONE,
		ActivationSignal := BUTTON_IMMEDIATE_STOP);

		// ON PHASE STOP
		SignalManagement
			(SignalType := ALARM,
			SignalCode := ID_ON_PHASE_STOP,
		SignalOutput := ON_PHASE_STOP OR NONE OR NONE,
		ActivationSignal := BUTTON_ON_PHASE_STOP);

		//######### FEEDER HANDLING SIGNALS #################//

		SignalManagement
		(SignalType := ALARM OR AUX_RESET,
		SignalCode := ID_CONVEYOR_IF_FAULT,
		SignalOutput := IMMEDIATE_STOP OR NONE OR NONE,
		ActivationSignal := CONVEYOR_IF_FAULT);

		SignalManagement
		(SignalType := ALARM OR AUX_RESET,
		SignalCode := ID_PUSHER_FAULT,
		SignalOutput := IMMEDIATE_STOP OR NONE OR NONE,
		ActivationSignal := PUSHER_FAULT);

		SignalManagement
		(SignalType := ALARM OR AUX_RESET,
		SignalCode := ID_TURNPUSHER_FAULT,
		SignalOutput := IMMEDIATE_STOP OR NONE OR NONE,
		ActivationSignal := TURNPUSHER_FAULT);

		SignalManagement
		(SignalType := ALARM OR AUX_RESET,
		SignalCode := ID_CONVEYOR_TURN1_FAULT,
		SignalOutput := IMMEDIATE_STOP OR NONE OR NONE,
		ActivationSignal := CONVEYOR_TURN1_FAULT);

		SignalManagement
		(SignalType := ALARM OR AUX_RESET,
		SignalCode := ID_CONVEYOR_END_FAULT,
		SignalOutput := IMMEDIATE_STOP OR NONE OR NONE,
		ActivationSignal := CONVEYOR_END_FAULT);

		SignalManagement
		(SignalType := ALARM OR AUX_RESET,
		SignalCode := ID_CARRIAGE_2_FAULT,
		SignalOutput := IMMEDIATE_STOP OR NONE OR NONE,
		ActivationSignal := CARRIAGE_2_FAULT);
		//######### CRANE HANDLING SIGNALS #################//
		SignalManagement
		(SignalType := ALARM OR AUX_RESET,
		SignalCode := ID_CARTBORAD_FAULT,
		SignalOutput := IMMEDIATE_STOP OR NONE OR NONE,
		ActivationSignal := CARTBORAD_FAULT);

		SignalManagement
		(SignalType := ALARM OR AUX_RESET,
		SignalCode := ID_VACUUM_BOX_CRANE_FAULT,
		SignalOutput := IMMEDIATE_STOP OR NONE OR NONE,
		ActivationSignal := VACUUM_BOX_CRANE_FAULT);

		SignalManagement
		(SignalType := ALARM OR AUX_RESET,
		SignalCode := ID_BOX_CRANE_FAULT,
		SignalOutput := IMMEDIATE_STOP OR NONE OR NONE,
		ActivationSignal := BOX_CRANE_FAULT);

		SignalManagement
		(SignalType := ALARM OR AUX_RESET,
		SignalCode := ID_GANTRY_CRANE_FAULT,
		SignalOutput := IMMEDIATE_STOP OR NONE OR NONE,
		ActivationSignal := GANTRY_CRANE_FAULT);

		SignalManagement
		(SignalType := ALARM OR AUX_RESET,
		SignalCode := ID_SLIDE_RAIL_RIGHT_FAULT,
		SignalOutput := IMMEDIATE_STOP OR NONE OR NONE,
		ActivationSignal := SLIDE_RAIL_RIGHT_FAULT);

		SignalManagement
		(SignalType := ALARM OR AUX_RESET,
		SignalCode := ID_PUSHER_X_FAULT,
		SignalOutput := IMMEDIATE_STOP OR NONE OR NONE,
		ActivationSignal := PUSHER_X_FAULT);

		SignalManagement
		(SignalType := ALARM OR AUX_RESET,
		SignalCode := ID_PUSHER_Z_FAULT,
		SignalOutput := IMMEDIATE_STOP OR NONE OR NONE,
		ActivationSignal := PUSHER_Z_FAULT);

							//######### PALLET HANDLING SIGNALS #################//
		IF PALLET_CONVEYOR_1_FAULT THEN
			coutn := coutn + 1;
		END_IF;
		SignalManagement
		(SignalType := ALARM OR AUX_RESET,
		SignalCode := ID_PALLET_CONVEYOR_1_FAULT,
		SignalOutput := IMMEDIATE_STOP OR NONE OR NONE,
		ActivationSignal := PALLET_CONVEYOR_1_FAULT );

		SignalManagement
		(SignalType := ALARM OR AUX_RESET,
		SignalCode := ID_PALLET_CONVEYOR_2_FAULT,
		SignalOutput := IMMEDIATE_STOP OR NONE OR NONE,
		ActivationSignal := PALLET_CONVEYOR_2_FAULT);

		SignalManagement
		(SignalType := ALARM OR AUX_RESET,
		SignalCode := ID_PALLET_LIFTER_FAULT,
		SignalOutput := IMMEDIATE_STOP OR NONE OR NONE,
		ActivationSignal := PALLET_LIFTER_FAULT);

		SignalManagement
		(SignalType := ALARM OR AUX_RESET,
		SignalCode := ID_PALLET_FORK_FAULT,
		SignalOutput := IMMEDIATE_STOP OR NONE OR NONE,
		ActivationSignal := PALLET_FORK_FAULT);

										//######### HANDLING SIGNAL OF CARTBOARD #################//

	END_IF;

	//######### OUTPUT HANDLING SIGNALS #################//
	CheckOperationSignals := SignalManagement.SignalOutputs;
	CathegorySIMSignalCode := SignalManagement.MySignalCode;
	Activate_signal			:= SignalManagement.ActiveSignalCodes;

	//######### VISUALISATION HANDLING SIGNALS GENRATION #################//
	IF (OperationType = RUN) THEN
		SignalManagement (OperationType := RUN); (* outputs selection *)
	END_IF;

	//############ PRIORYTY MANAGEMENT OF SIGNALS ##################### //
	SM_EMERGENCY_STOP := ((CheckOperationSignals AND EMERGENCY_STOP) = EMERGENCY_STOP);

	IF SM_EMERGENCY_STOP  THEN
		SM_IMMEDIATE_STOP		:= FALSE;
		SM_IMMEDIATE_STOP_CAT1	:= FALSE;
		SM_IMMEDIATE_STOP_CAT2	:= FALSE;
		SM_IMMEDIATE_STOP_CAT3	:= FALSE;
		SM_ON_PHASE_STOP 		:= FALSE;
		blink_emergencvy_stop 	:= NOT blink_emergencvy_stop;
	END_IF;

	IF NOT SM_EMERGENCY_STOP  THEN
		blink_emergencvy_stop 	:= FALSE;
		IF CathegorySIMSignalCode = 2 THEN
			blink_immediate_stop 	:= NOT blink_immediate_stop;

			SM_IMMEDIATE_STOP := ((CheckOperationSignals AND IMMEDIATE_STOP) = IMMEDIATE_STOP);
			SM_IMMEDIATE_STOP_CAT1	:= FALSE;
		END_IF;
		IF  CathegorySIMSignalCode>3 AND CathegorySIMSignalCode<=20 AND NOT SM_IMMEDIATE_STOP THEN
			blink_immediate_stop 	:= NOT blink_immediate_stop;
			SM_IMMEDIATE_STOP_CAT1  := ((CheckOperationSignals AND IMMEDIATE_STOP) = IMMEDIATE_STOP);
		END_IF;

		IF SM_IMMEDIATE_STOP_CAT1 OR SM_IMMEDIATE_STOP THEN
			SM_ON_PHASE_STOP	:= FALSE;
			SM_ON_PHASE_STOP_CAT1	:= FALSE;
			SM_ON_PHASE_STOP_CAT2	:= FALSE;
		END_IF;
	END_IF;

	IF NOT SM_IMMEDIATE_STOP_CAT1 AND  NOT SM_IMMEDIATE_STOP  THEN
		blink_immediate_stop 	:= FALSE;
		IF (CathegorySIMSignalCode =3) THEN
			blink_OnPhase_stop 	:= NOT blink_OnPhase_stop;
			SM_ON_PHASE_STOP  := ((CheckOperationSignals AND ON_PHASE_STOP) = ON_PHASE_STOP);
			SM_ON_PHASE_STOP_CAT1	:= FALSE;
		END_IF
		IF  (CathegorySIMSignalCode =22) AND NOT SM_ON_PHASE_STOP  THEN
			blink_OnPhase_stop 	:= NOT blink_OnPhase_stop;
			SM_ON_PHASE_STOP_CAT1  := ((CheckOperationSignals AND ON_PHASE_STOP) = ON_PHASE_STOP);
		END_IF;
		IF NOT SM_ON_PHASE_STOP_CAT1 AND NOT SM_ON_PHASE_STOP THEN
			blink_OnPhase_stop 	:= FALSE;
		END_IF;
	END_IF;

	LED_MATERIALS_RUN_OUT	:= ((CheckOperationSignals AND MATERIALS_RUN_OUT_LAMP) = MATERIALS_RUN_OUT_LAMP);

	LED_ALARM_INFORMATION := SignalManagement.LedSignalInformation;
	LED_ALARM_ANOMALY := SignalManagement.LedSignalAnomaly;
	LED_ALARM_ALARM := SignalManagement.LedSignalAlarm ;
	LED_ALARM_WARNING := SignalManagement.LedSignalWarning;
	IF pallet_lifter_ALMOST_FINISH OR boxcrane_Cartboard_ALMOST_FINISH THEN
		blink_out_of_material:=TRUE;
	ELSE
		blink_out_of_material:=FALSE;
	END_IF;

END_PROGRAM

PROGRAM _EXIT
	(* Insert code here *)

END_PROGRAM
```

#### Variables.var - Local variables
```iecst
VAR
	SignalManagement : GenericSignalHandler;
	CheckOperationSignals : DWORD;
	CathegorySIMSignalCode : INT;
END_VAR
VAR CONSTANT
	ID_EMERGENCY_STOP : INT := 1;
	ID_IMMEDIATE_STOP : INT := 2;
	ID_ON_PHASE_STOP : INT := 3;
	ID_CONVEYOR_IF_FAULT : INT := 4;
	ID_PUSHER_FAULT : INT := 5;
	ID_TURNPUSHER_FAULT : INT := 6;
	ID_CONVEYOR_TURN1_FAULT : INT := 7;
	ID_CONVEYOR_END_FAULT : INT := 8;
	ID_CARRIAGE_2_FAULT : INT := 9;
	ID_CARTBORAD_FAULT : INT := 10;
	ID_VACUUM_BOX_CRANE_FAULT : INT := 11;
	ID_BOX_CRANE_FAULT : INT := 12;
	ID_GANTRY_CRANE_FAULT : INT := 13;
	ID_SLIDE_RAIL_RIGHT_FAULT : INT := 14;
	ID_PUSHER_X_FAULT : INT := 15;
	ID_PUSHER_Z_FAULT : INT := 16;
	ID_PALLET_CONVEYOR_1_FAULT : INT := 17;
	ID_PALLET_CONVEYOR_2_FAULT : INT := 18;
	ID_PALLET_LIFTER_FAULT : INT := 19;
	ID_PALLET_FORK_FAULT : INT := 20;
	ID_Cartboard_ALMOST_FINISH : INT := 21;
	ID_Cartboard_FINISH : INT := 22;
	ID_P_lifter_ALMOST_FINISH : INT := 23;
	ID_pallet_lifter_FINISH : INT := 24;
END_VAR
VAR
	Activate_signal : ARRAY[0..24] OF INT;
	PALLET_CONVEYOR_1_FAULT_my : BOOL;
	CountEnablingTimer : BOOL := FALSE;
	Count : INT := 600;
	coutn : INT;
	blink_out_of_material : BOOL;
END_VAR
```

### MNG_Global.typ - Global data types
```iecst
(* 3d position *)
(* position and orientation as an euler based pose *)
(* position and orientation as a 4x4 matrix *)

TYPE
	VEC3 : 	STRUCT
		x : REAL;
		y : REAL;
		z : REAL;
	END_STRUCT;
	POSE6 : 	STRUCT
		x : REAL;
		y : REAL;
		z : REAL;
		a : REAL;
		b : REAL;
		c : REAL;
	END_STRUCT;
	TRAFO : 	STRUCT
		baseX : VEC3;
		fill0 : REAL;
		baseY : VEC3;
		fill1 : REAL;
		baseZ : VEC3;
		fill2 : REAL;
		origin : VEC3;
		fill3 : REAL;
	END_STRUCT;
END_TYPE
```

- Visualisation Logical/Visu_Resized (not shown)

Listed in the project but not available here: Logical/Libraries/ComTCP
